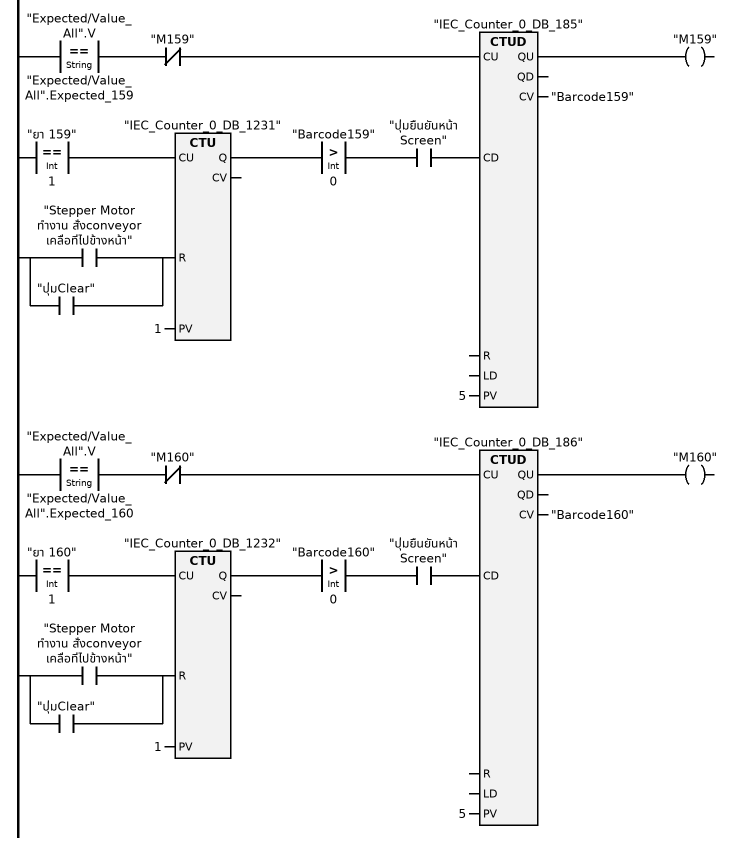
   "IEC_Counter_0_DB_1213".CTU(CU := "ยา 141" = 1,
                           R := "Stepper Motor ทำงาน สั่งconveyor เคลื่อที่ไปข้างหน้า" OR "ปุ่มClear",
                           PV := 1);
   "IEC_Counter_0_DB_167".CTUD(CU := ("Expected/Value_All".V = "Expected/Value_All".Expected_141) AND NOT "M141",
                           CD := "IEC_Counter_0_DB_1213".Q AND ("Barcode141" > 0) AND "ปุ่มยืนยันหน้า Screen",
                           PV := 5,
                           CV => "Barcode141");
   "M141" := "IEC_Counter_0_DB_167".QU;
   "IEC_Counter_0_DB_1214".CTU(CU := "ยา 142" = 1,
                           R := "Stepper Motor ทำงาน สั่งconveyor เคลื่อที่ไปข้างหน้า" OR "ปุ่มClear",
                           PV := 1);
   "IEC_Counter_0_DB_168".CTUD(CU := ("Expected/Value_All".V = "Expected/Value_All".Expected_142) AND NOT "M142",
                           CD := "IEC_Counter_0_DB_1214".Q AND ("Barcode142" > 0) AND "ปุ่มยืนยันหน้า Screen",
                           PV := 5,
                           CV => "Barcode142");
   "M142" := "IEC_Counter_0_DB_168".QU;
   "IEC_Counter_0_DB_1215".CTU(CU := "ยา 143" = 1,
                           R := "Stepper Motor ทำงาน สั่งconveyor เคลื่อที่ไปข้างหน้า" OR "ปุ่มClear",
                           PV := 1);
   "IEC_Counter_0_DB_169".CTUD(CU := ("Expected/Value_All".V = "Expected/Value_All".Expected_143) AND NOT "M143",
                           CD := "IEC_Counter_0_DB_1215".Q AND ("Barcode143" > 0) AND "ปุ่มยืนยันหน้า Screen",
                           PV := 5,
                           CV => "Barcode143");
   "M143" := "IEC_Counter_0_DB_169".QU;
   "IEC_Counter_0_DB_1216".CTU(CU := "ยา 144" = 1,
                           R := "Stepper Motor ทำงาน สั่งconveyor เคลื่อที่ไปข้างหน้า" OR "ปุ่มClear",
                           PV := 1);
   "IEC_Counter_0_DB_170".CTUD(CU := ("Expected/Value_All".V = "Expected/Value_All".Expected_144) AND NOT "M144",
                           CD := "IEC_Counter_0_DB_1216".Q AND ("Barcode144" > 0) AND "ปุ่มยืนยันหน้า Screen",
                           PV := 5,
                           CV => "Barcode144");
   "M144" := "IEC_Counter_0_DB_170".QU;
   "IEC_Counter_0_DB_1217".CTU(CU := "ยา 145" = 1,
                           R := "Stepper Motor ทำงาน สั่งconveyor เคลื่อที่ไปข้างหน้า" OR "ปุ่มClear",
                           PV := 1);
   "IEC_Counter_0_DB_171".CTUD(CU := ("Expected/Value_All".V = "Expected/Value_All".Expected_145) AND NOT "M145",
                           CD := "IEC_Counter_0_DB_1217".Q AND ("Barcode145" > 0) AND "ปุ่มยืนยันหน้า Screen",
                           PV := 5,
                           CV => "Barcode145");
   "M145" := "IEC_Counter_0_DB_171".QU;
   "IEC_Counter_0_DB_1218".CTU(CU := "ยา 146" = 1,
                           R := "Stepper Motor ทำงาน สั่งconveyor เคลื่อที่ไปข้างหน้า" OR "ปุ่มClear",
                           PV := 1);
   "IEC_Counter_0_DB_172".CTUD(CU := ("Expected/Value_All".V = "Expected/Value_All".Expected_146) AND NOT "M146",
                           CD := "IEC_Counter_0_DB_1218".Q AND ("Barcode146" > 0) AND "ปุ่มยืนยันหน้า Screen",
                           PV := 5,
                           CV => "Barcode146");
   "M146" := "IEC_Counter_0_DB_172".QU;
   "IEC_Counter_0_DB_1219".CTU(CU := "ยา 147" = 1,
                           R := "Stepper Motor ทำงาน สั่งconveyor เคลื่อที่ไปข้างหน้า" OR "ปุ่มClear",
                           PV := 1);
   "IEC_Counter_0_DB_173".CTUD(CU := ("Expected/Value_All".V = "Expected/Value_All".Expected_147) AND NOT "M147",
                           CD := "IEC_Counter_0_DB_1219".Q AND ("Barcode147" > 0) AND "ปุ่มยืนยันหน้า Screen",
                           PV := 5,
                           CV => "Barcode147");
   "M147" := "IEC_Counter_0_DB_173".QU;
   "IEC_Counter_0_DB_1220".CTU(CU := "ยา 148" = 1,
                           R := "Stepper Motor ทำงาน สั่งconveyor เคลื่อที่ไปข้างหน้า" OR "ปุ่มClear",
                           PV := 1);
   "IEC_Counter_0_DB_174".CTUD(CU := ("Expected/Value_All".V = "Expected/Value_All".Expected_148) AND NOT "M148",
                           CD := "IEC_Counter_0_DB_1220".Q AND ("Barcode148" > 0) AND "ปุ่มยืนยันหน้า Screen",
                           PV := 5,
                           CV => "Barcode148");
   "M148" := "IEC_Counter_0_DB_174".QU;
   "IEC_Counter_0_DB_1221".CTU(CU := "ยา 149" = 1,
                           R := "Stepper Motor ทำงาน สั่งconveyor เคลื่อที่ไปข้างหน้า" OR "ปุ่มClear",
                           PV := 1);
   "IEC_Counter_0_DB_175".CTUD(CU := ("Expected/Value_All".V = "Expected/Value_All".Expected_149) AND NOT "M149",
                           CD := "IEC_Counter_0_DB_1221".Q AND ("Barcode149" > 0) AND "ปุ่มยืนยันหน้า Screen",
                           PV := 5,
                           CV => "Barcode149");
   "M149" := "IEC_Counter_0_DB_175".QU;
   "IEC_Counter_0_DB_1222".CTU(CU := "ยา 150" = 1,
                           R := "Stepper Motor ทำงาน สั่งconveyor เคลื่อที่ไปข้างหน้า" OR "ปุ่มClear",
                           PV := 1);
   "IEC_Counter_0_DB_176".CTUD(CU := ("Expected/Value_All".V = "Expected/Value_All".Expected_150) AND NOT "M150",
                           CD := "IEC_Counter_0_DB_1222".Q AND ("Barcode150" > 0) AND "ปุ่มยืนยันหน้า Screen",
                           PV := 5,
                           CV => "Barcode150");
   "M150" := "IEC_Counter_0_DB_176".QU;
   "IEC_Counter_0_DB_1223".CTU(CU := "ยา 151" = 1,
                           R := "Stepper Motor ทำงาน สั่งconveyor เคลื่อที่ไปข้างหน้า" OR "ปุ่มClear",
                           PV := 1);
   "IEC_Counter_0_DB_177".CTUD(CU := ("Expected/Value_All".V = "Expected/Value_All".Expected_151) AND NOT "M151",
                           CD := "IEC_Counter_0_DB_1223".Q AND ("Barcode151" > 0) AND "ปุ่มยืนยันหน้า Screen",
                           PV := 5,
                           CV => "Barcode151");
   "M151" := "IEC_Counter_0_DB_177".QU;
   "IEC_Counter_0_DB_1224".CTU(CU := "ยา 152" = 1,
                           R := "Stepper Motor ทำงาน สั่งconveyor เคลื่อที่ไปข้างหน้า" OR "ปุ่มClear",
                           PV := 1);
   "IEC_Counter_0_DB_178".CTUD(CU := ("Expected/Value_All".V = "Expected/Value_All".Expected_152) AND NOT "M152",
                           CD := "IEC_Counter_0_DB_1224".Q AND ("Barcode152" > 0) AND "ปุ่มยืนยันหน้า Screen",
                           PV := 5,
                           CV => "Barcode152");
   "M152" := "IEC_Counter_0_DB_178".QU;
   "IEC_Counter_0_DB_1225".CTU(CU := "ยา 153" = 1,
                           R := "Stepper Motor ทำงาน สั่งconveyor เคลื่อที่ไปข้างหน้า" OR "ปุ่มClear",
                           PV := 1);
   "IEC_Counter_0_DB_179".CTUD(CU := ("Expected/Value_All".V = "Expected/Value_All".Expected_153) AND NOT "M153",
                           CD := "IEC_Counter_0_DB_1225".Q AND ("Barcode153" > 0) AND "ปุ่มยืนยันหน้า Screen",
                           PV := 5,
                           CV => "Barcode153");
   "M153" := "IEC_Counter_0_DB_179".QU;
   "IEC_Counter_0_DB_1226".CTU(CU := "ยา 154" = 1,
                           R := "Stepper Motor ทำงาน สั่งconveyor เคลื่อที่ไปข้างหน้า" OR "ปุ่มClear",
                           PV := 1);
   "IEC_Counter_0_DB_180".CTUD(CU := ("Expected/Value_All".V = "Expected/Value_All".Expected_154) AND NOT "M154",
                           CD := "IEC_Counter_0_DB_1226".Q AND ("Barcode154" > 0) AND "ปุ่มยืนยันหน้า Screen",
                           PV := 5,
                           CV => "Barcode154");
   "M154" := "IEC_Counter_0_DB_180".QU;
   "IEC_Counter_0_DB_1227".CTU(CU := "ยา 155" = 1,
                           R := "Stepper Motor ทำงาน สั่งconveyor เคลื่อที่ไปข้างหน้า" OR "ปุ่มClear",
                           PV := 1);
   "IEC_Counter_0_DB_181".CTUD(CU := ("Expected/Value_All".V = "Expected/Value_All".Expected_155) AND NOT "M155",
                           CD := "IEC_Counter_0_DB_1227".Q AND ("Barcode155" > 0) AND "ปุ่มยืนยันหน้า Screen",
                           PV := 5,
                           CV => "Barcode155");
   "M155" := "IEC_Counter_0_DB_181".QU;
   "IEC_Counter_0_DB_1228".CTU(CU := "ยา 156" = 1,
                           R := "Stepper Motor ทำงาน สั่งconveyor เคลื่อที่ไปข้างหน้า" OR "ปุ่มClear",
                           PV := 1);
   "IEC_Counter_0_DB_182".CTUD(CU := ("Expected/Value_All".V = "Expected/Value_All".Expected_156) AND NOT "M156",
                           CD := "IEC_Counter_0_DB_1228".Q AND ("Barcode156" > 0) AND "ปุ่มยืนยันหน้า Screen",
                           PV := 5,
                           CV => "Barcode156");
   "M156" := "IEC_Counter_0_DB_182".QU;
   "IEC_Counter_0_DB_1229".CTU(CU := "ยา 157" = 1,
                           R := "Stepper Motor ทำงาน สั่งconveyor เคลื่อที่ไปข้างหน้า" OR "ปุ่มClear",
                           PV := 1);
   "IEC_Counter_0_DB_183".CTUD(CU := ("Expected/Value_All".V = "Expected/Value_All".Expected_157) AND NOT "M157",
                           CD := "IEC_Counter_0_DB_1229".Q AND ("Barcode157" > 0) AND "ปุ่มยืนยันหน้า Screen",
                           PV := 5,
                           CV => "Barcode157");
   "M157" := "IEC_Counter_0_DB_183".QU;
   "IEC_Counter_0_DB_1230".CTU(CU := "ยา 158" = 1,
                           R := "Stepper Motor ทำงาน สั่งconveyor เคลื่อที่ไปข้างหน้า" OR "ปุ่มClear",
                           PV := 1);
   "IEC_Counter_0_DB_184".CTUD(CU := ("Expected/Value_All".V = "Expected/Value_All".Expected_158) AND NOT "M158",
                           CD := "IEC_Counter_0_DB_1230".Q AND ("Barcode158" > 0) AND "ปุ่มยืนยันหน้า Screen",
                           PV := 5,
                           CV => "Barcode158");
   "M158" := "IEC_Counter_0_DB_184".QU;
   "IEC_Counter_0_DB_1231".CTU(CU := "ยา 159" = 1,
                           R := "Stepper Motor ทำงาน สั่งconveyor เคลื่อที่ไปข้างหน้า" OR "ปุ่มClear",
                           PV := 1);
   "IEC_Counter_0_DB_185".CTUD(CU := ("Expected/Value_All".V = "Expected/Value_All".Expected_159) AND NOT "M159",
                           CD := "IEC_Counter_0_DB_1231".Q AND ("Barcode159" > 0) AND "ปุ่มยืนยันหน้า Screen",
                           PV := 5,
                           CV => "Barcode159");
   "M159" := "IEC_Counter_0_DB_185".QU;
   "IEC_Counter_0_DB_1232".CTU(CU := "ยา 160" = 1,
                           R := "Stepper Motor ทำงาน สั่งconveyor เคลื่อที่ไปข้างหน้า" OR "ปุ่มClear",
                           PV := 1);
   "IEC_Counter_0_DB_186".CTUD(CU := ("Expected/Value_All".V = "Expected/Value_All".Expected_160) AND NOT "M160",
                           CD := "IEC_Counter_0_DB_1232".Q AND ("Barcode160" > 0) AND "ปุ่มยืนยันหน้า Screen",
                           PV := 5,
                           CV => "Barcode160");
   "M160" := "IEC_Counter_0_DB_186".QU;
END_REGION

REGION Network 9
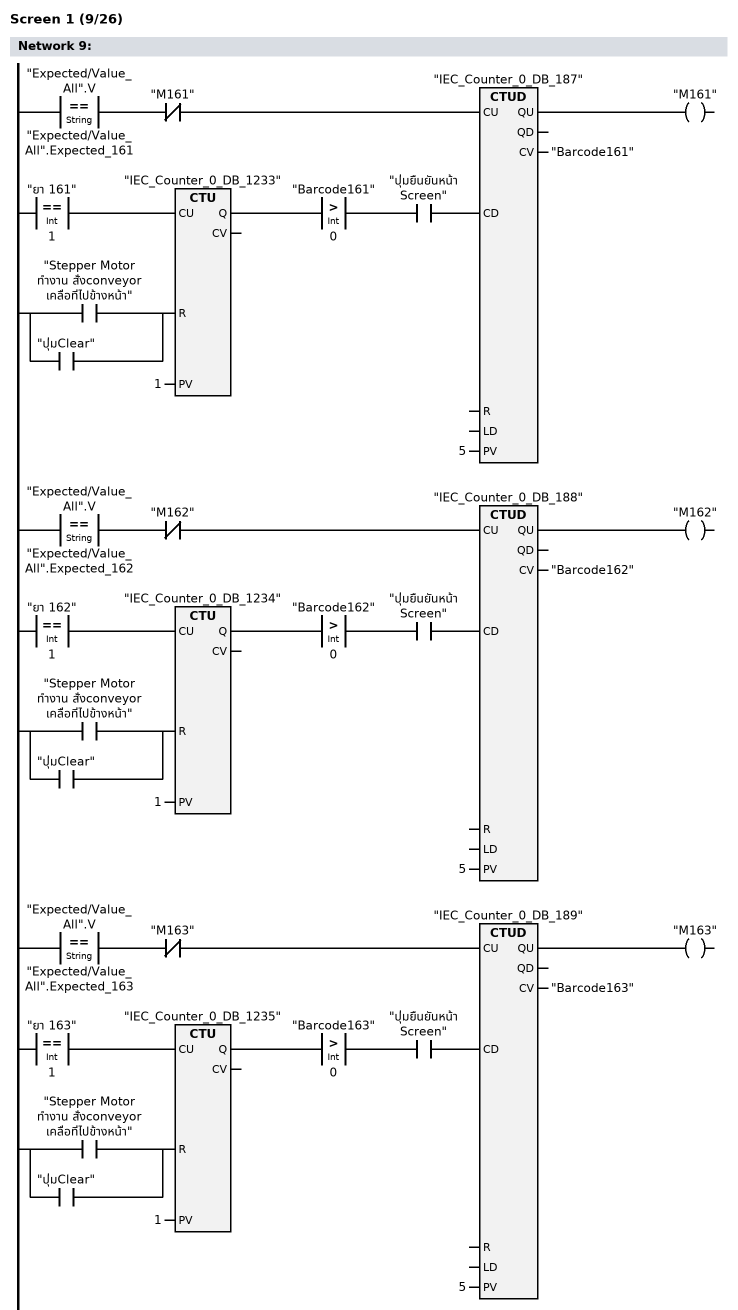
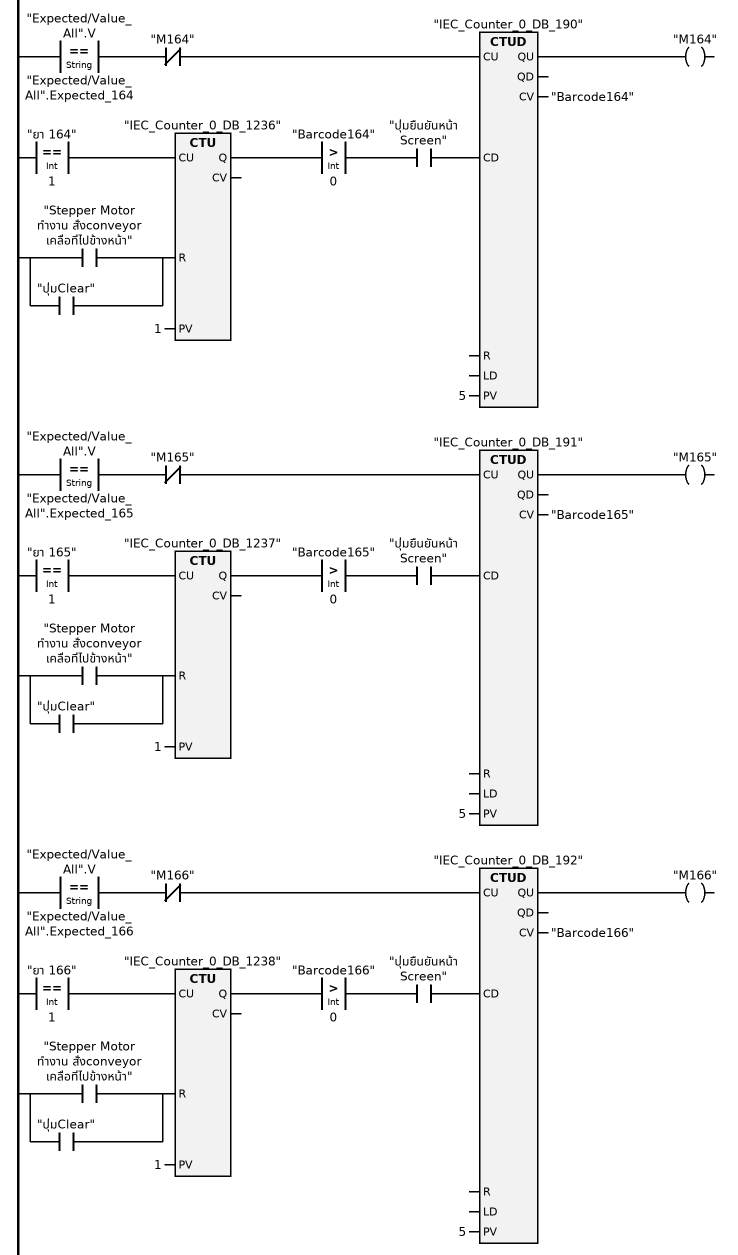
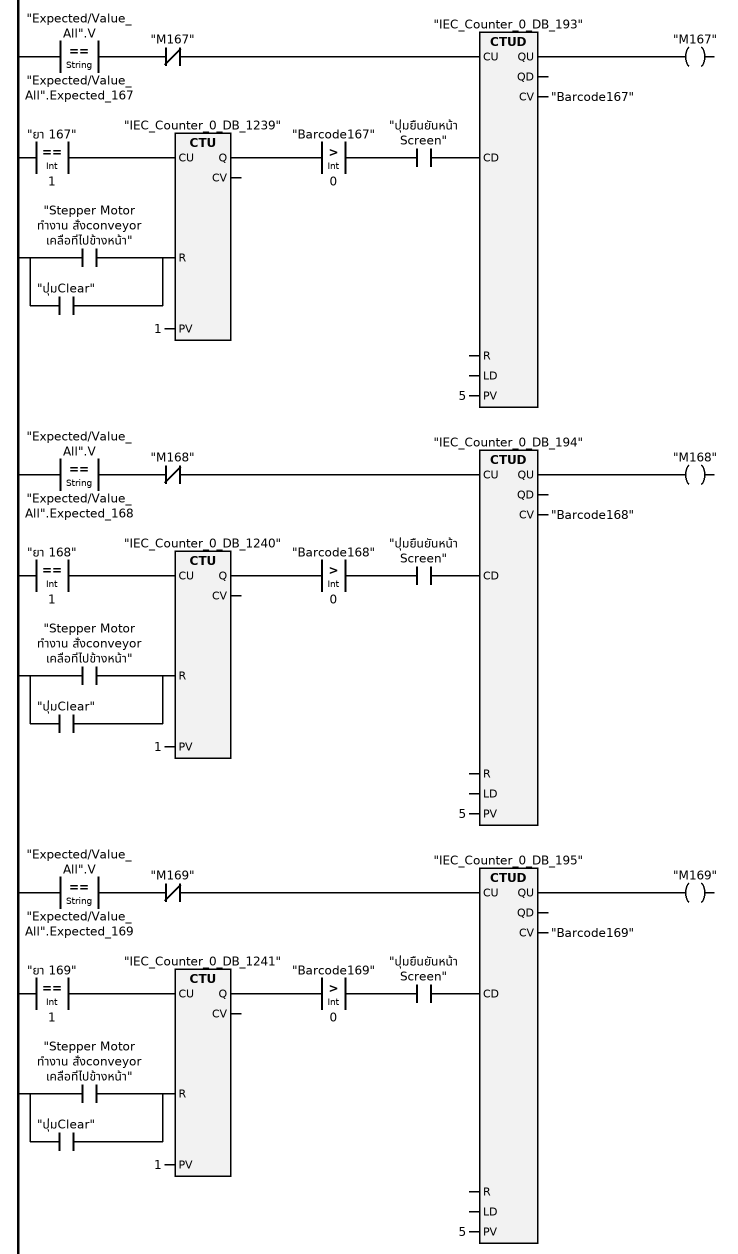
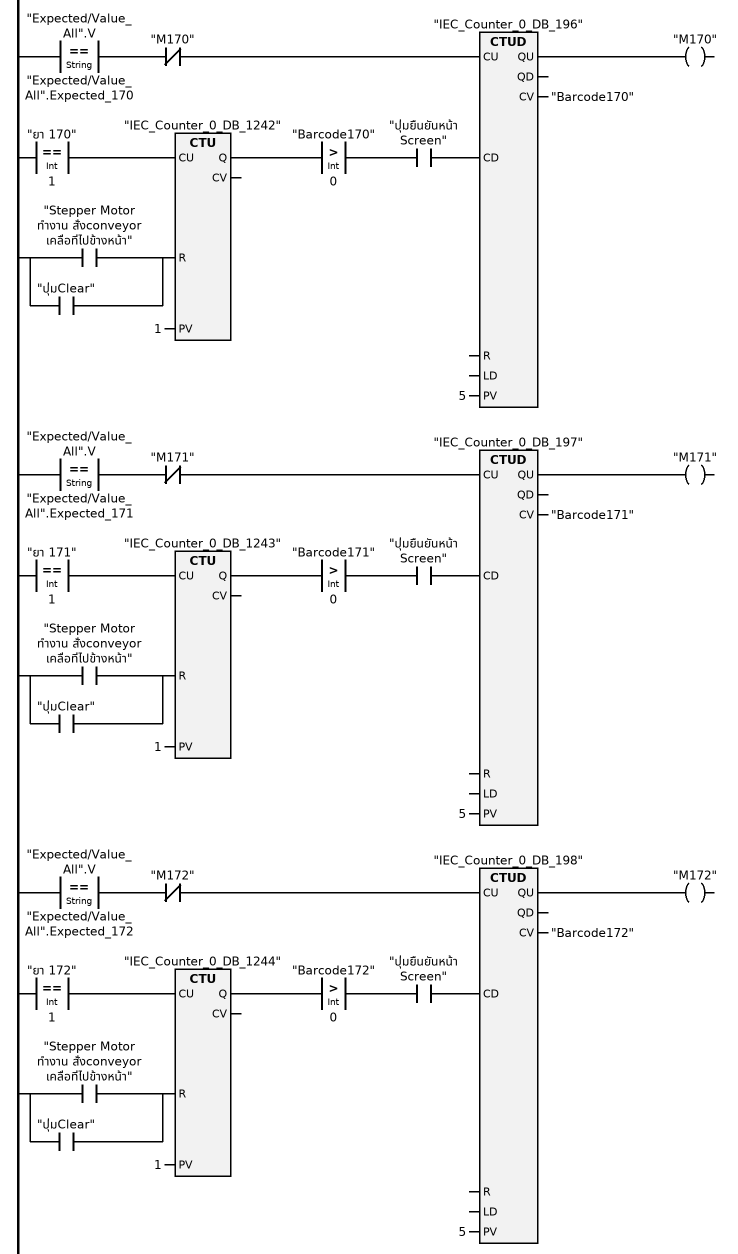
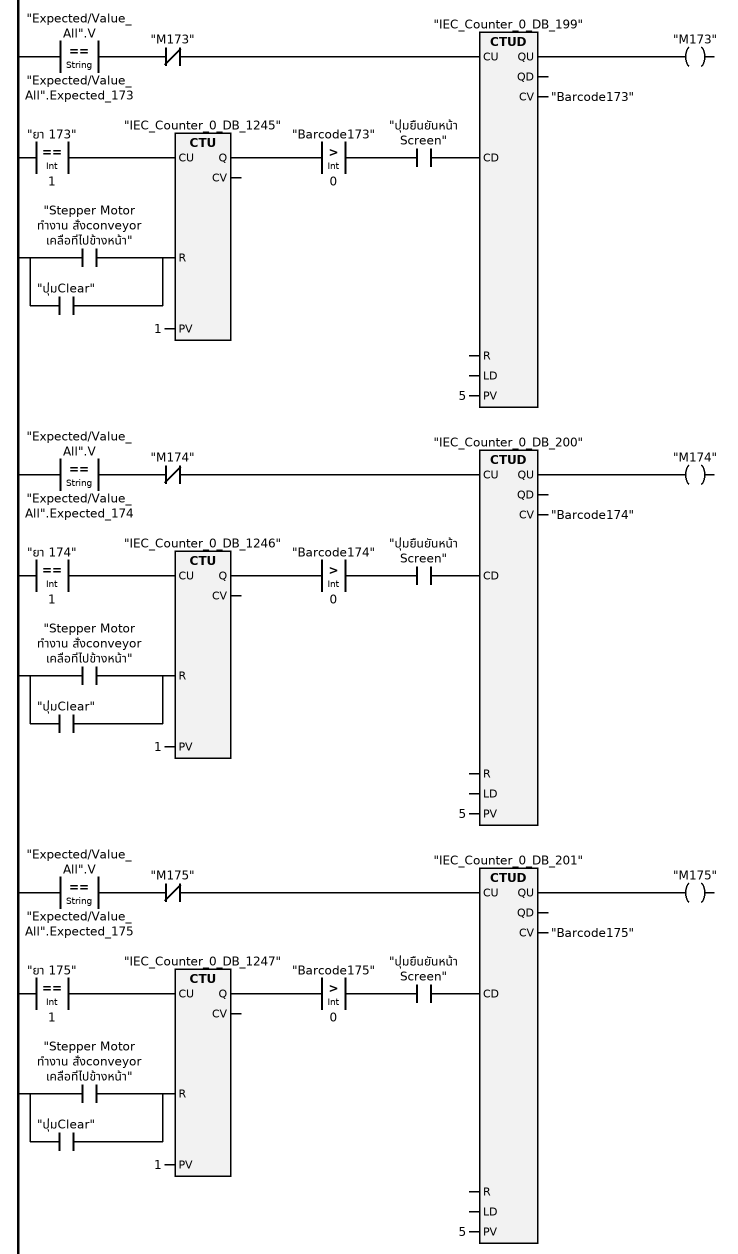
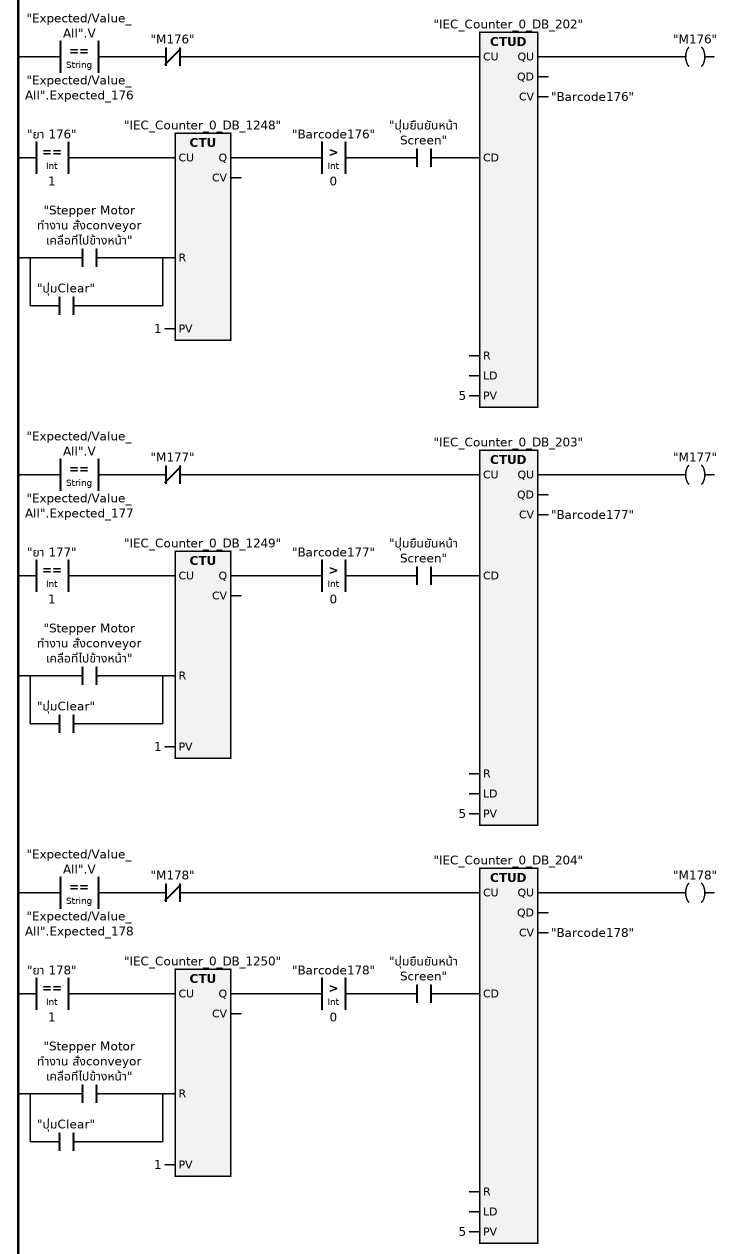
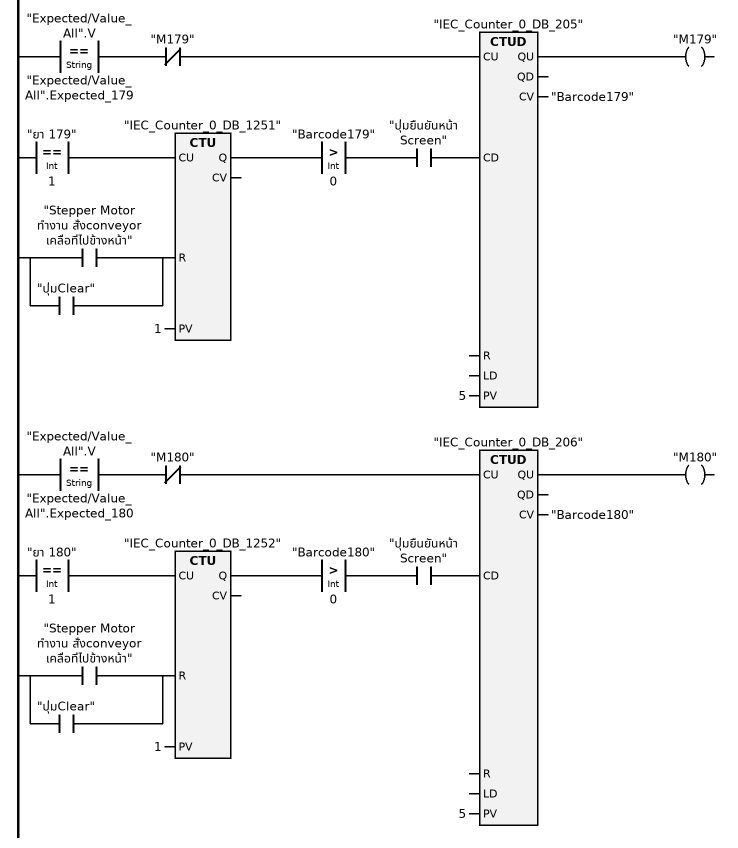
   "IEC_Counter_0_DB_1233".CTU(CU := "ยา 161" = 1,
                           R := "Stepper Motor ทำงาน สั่งconveyor เคลื่อที่ไปข้างหน้า" OR "ปุ่มClear",
                           PV := 1);
   "IEC_Counter_0_DB_187".CTUD(CU := ("Expected/Value_All".V = "Expected/Value_All".Expected_161) AND NOT "M161",
                           CD := "IEC_Counter_0_DB_1233".Q AND ("Barcode161" > 0) AND "ปุ่มยืนยันหน้า Screen",
                           PV := 5,
                           CV => "Barcode161");
   "M161" := "IEC_Counter_0_DB_187".QU;
   "IEC_Counter_0_DB_1234".CTU(CU := "ยา 162" = 1,
                           R := "Stepper Motor ทำงาน สั่งconveyor เคลื่อที่ไปข้างหน้า" OR "ปุ่มClear",
                           PV := 1);
   "IEC_Counter_0_DB_188".CTUD(CU := ("Expected/Value_All".V = "Expected/Value_All".Expected_162) AND NOT "M162",
                           CD := "IEC_Counter_0_DB_1234".Q AND ("Barcode162" > 0) AND "ปุ่มยืนยันหน้า Screen",
                           PV := 5,
                           CV => "Barcode162");
   "M162" := "IEC_Counter_0_DB_188".QU;
   "IEC_Counter_0_DB_1235".CTU(CU := "ยา 163" = 1,
                           R := "Stepper Motor ทำงาน สั่งconveyor เคลื่อที่ไปข้างหน้า" OR "ปุ่มClear",
                           PV := 1);
   "IEC_Counter_0_DB_189".CTUD(CU := ("Expected/Value_All".V = "Expected/Value_All".Expected_163) AND NOT "M163",
                           CD := "IEC_Counter_0_DB_1235".Q AND ("Barcode163" > 0) AND "ปุ่มยืนยันหน้า Screen",
                           PV := 5,
                           CV => "Barcode163");
   "M163" := "IEC_Counter_0_DB_189".QU;
   "IEC_Counter_0_DB_1236".CTU(CU := "ยา 164" = 1,
                           R := "Stepper Motor ทำงาน สั่งconveyor เคลื่อที่ไปข้างหน้า" OR "ปุ่มClear",
                           PV := 1);
   "IEC_Counter_0_DB_190".CTUD(CU := ("Expected/Value_All".V = "Expected/Value_All".Expected_164) AND NOT "M164",
                           CD := "IEC_Counter_0_DB_1236".Q AND ("Barcode164" > 0) AND "ปุ่มยืนยันหน้า Screen",
                           PV := 5,
                           CV => "Barcode164");
   "M164" := "IEC_Counter_0_DB_190".QU;
   "IEC_Counter_0_DB_1237".CTU(CU := "ยา 165" = 1,
                           R := "Stepper Motor ทำงาน สั่งconveyor เคลื่อที่ไปข้างหน้า" OR "ปุ่มClear",
                           PV := 1);
   "IEC_Counter_0_DB_191".CTUD(CU := ("Expected/Value_All".V = "Expected/Value_All".Expected_165) AND NOT "M165",
                           CD := "IEC_Counter_0_DB_1237".Q AND ("Barcode165" > 0) AND "ปุ่มยืนยันหน้า Screen",
                           PV := 5,
                           CV => "Barcode165");
   "M165" := "IEC_Counter_0_DB_191".QU;
   "IEC_Counter_0_DB_1238".CTU(CU := "ยา 166" = 1,
                           R := "Stepper Motor ทำงาน สั่งconveyor เคลื่อที่ไปข้างหน้า" OR "ปุ่มClear",
                           PV := 1);
   "IEC_Counter_0_DB_192".CTUD(CU := ("Expected/Value_All".V = "Expected/Value_All".Expected_166) AND NOT "M166",
                           CD := "IEC_Counter_0_DB_1238".Q AND ("Barcode166" > 0) AND "ปุ่มยืนยันหน้า Screen",
                           PV := 5,
                           CV => "Barcode166");
   "M166" := "IEC_Counter_0_DB_192".QU;
   "IEC_Counter_0_DB_1239".CTU(CU := "ยา 167" = 1,
                           R := "Stepper Motor ทำงาน สั่งconveyor เคลื่อที่ไปข้างหน้า" OR "ปุ่มClear",
                           PV := 1);
   "IEC_Counter_0_DB_193".CTUD(CU := ("Expected/Value_All".V = "Expected/Value_All".Expected_167) AND NOT "M167",
                           CD := "IEC_Counter_0_DB_1239".Q AND ("Barcode167" > 0) AND "ปุ่มยืนยันหน้า Screen",
                           PV := 5,
                           CV => "Barcode167");
   "M167" := "IEC_Counter_0_DB_193".QU;
   "IEC_Counter_0_DB_1240".CTU(CU := "ยา 168" = 1,
                           R := "Stepper Motor ทำงาน สั่งconveyor เคลื่อที่ไปข้างหน้า" OR "ปุ่มClear",
                           PV := 1);
   "IEC_Counter_0_DB_194".CTUD(CU := ("Expected/Value_All".V = "Expected/Value_All".Expected_168) AND NOT "M168",
                           CD := "IEC_Counter_0_DB_1240".Q AND ("Barcode168" > 0) AND "ปุ่มยืนยันหน้า Screen",
                           PV := 5,
                           CV => "Barcode168");
   "M168" := "IEC_Counter_0_DB_194".QU;
   "IEC_Counter_0_DB_1241".CTU(CU := "ยา 169" = 1,
                           R := "Stepper Motor ทำงาน สั่งconveyor เคลื่อที่ไปข้างหน้า" OR "ปุ่มClear",
                           PV := 1);
   "IEC_Counter_0_DB_195".CTUD(CU := ("Expected/Value_All".V = "Expected/Value_All".Expected_169) AND NOT "M169",
                           CD := "IEC_Counter_0_DB_1241".Q AND ("Barcode169" > 0) AND "ปุ่มยืนยันหน้า Screen",
                           PV := 5,
                           CV => "Barcode169");
   "M169" := "IEC_Counter_0_DB_195".QU;
   "IEC_Counter_0_DB_1242".CTU(CU := "ยา 170" = 1,
                           R := "Stepper Motor ทำงาน สั่งconveyor เคลื่อที่ไปข้างหน้า" OR "ปุ่มClear",
                           PV := 1);
   "IEC_Counter_0_DB_196".CTUD(CU := ("Expected/Value_All".V = "Expected/Value_All".Expected_170) AND NOT "M170",
                           CD := "IEC_Counter_0_DB_1242".Q AND ("Barcode170" > 0) AND "ปุ่มยืนยันหน้า Screen",
                           PV := 5,
                           CV => "Barcode170");
   "M170" := "IEC_Counter_0_DB_196".QU;
   "IEC_Counter_0_DB_1243".CTU(CU := "ยา 171" = 1,
                           R := "Stepper Motor ทำงาน สั่งconveyor เคลื่อที่ไปข้างหน้า" OR "ปุ่มClear",
                           PV := 1);
   "IEC_Counter_0_DB_197".CTUD(CU := ("Expected/Value_All".V = "Expected/Value_All".Expected_171) AND NOT "M171",
                           CD := "IEC_Counter_0_DB_1243".Q AND ("Barcode171" > 0) AND "ปุ่มยืนยันหน้า Screen",
                           PV := 5,
                           CV => "Barcode171");
   "M171" := "IEC_Counter_0_DB_197".QU;
   "IEC_Counter_0_DB_1244".CTU(CU := "ยา 172" = 1,
                           R := "Stepper Motor ทำงาน สั่งconveyor เคลื่อที่ไปข้างหน้า" OR "ปุ่มClear",
                           PV := 1);
   "IEC_Counter_0_DB_198".CTUD(CU := ("Expected/Value_All".V = "Expected/Value_All".Expected_172) AND NOT "M172",
                           CD := "IEC_Counter_0_DB_1244".Q AND ("Barcode172" > 0) AND "ปุ่มยืนยันหน้า Screen",
                           PV := 5,
                           CV => "Barcode172");
   "M172" := "IEC_Counter_0_DB_198".QU;
   "IEC_Counter_0_DB_1245".CTU(CU := "ยา 173" = 1,
                           R := "Stepper Motor ทำงาน สั่งconveyor เคลื่อที่ไปข้างหน้า" OR "ปุ่มClear",
                           PV := 1);
   "IEC_Counter_0_DB_199".CTUD(CU := ("Expected/Value_All".V = "Expected/Value_All".Expected_173) AND NOT "M173",
                           CD := "IEC_Counter_0_DB_1245".Q AND ("Barcode173" > 0) AND "ปุ่มยืนยันหน้า Screen",
                           PV := 5,
                           CV => "Barcode173");
   "M173" := "IEC_Counter_0_DB_199".QU;
   "IEC_Counter_0_DB_1246".CTU(CU := "ยา 174" = 1,
                           R := "Stepper Motor ทำงาน สั่งconveyor เคลื่อที่ไปข้างหน้า" OR "ปุ่มClear",
                           PV := 1);
   "IEC_Counter_0_DB_200".CTUD(CU := ("Expected/Value_All".V = "Expected/Value_All".Expected_174) AND NOT "M174",
                           CD := "IEC_Counter_0_DB_1246".Q AND ("Barcode174" > 0) AND "ปุ่มยืนยันหน้า Screen",
                           PV := 5,
                           CV => "Barcode174");
   "M174" := "IEC_Counter_0_DB_200".QU;
   "IEC_Counter_0_DB_1247".CTU(CU := "ยา 175" = 1,
                           R := "Stepper Motor ทำงาน สั่งconveyor เคลื่อที่ไปข้างหน้า" OR "ปุ่มClear",
                           PV := 1);
   "IEC_Counter_0_DB_201".CTUD(CU := ("Expected/Value_All".V = "Expected/Value_All".Expected_175) AND NOT "M175",
                           CD := "IEC_Counter_0_DB_1247".Q AND ("Barcode175" > 0) AND "ปุ่มยืนยันหน้า Screen",
                           PV := 5,
                           CV => "Barcode175");
   "M175" := "IEC_Counter_0_DB_201".QU;
   "IEC_Counter_0_DB_1248".CTU(CU := "ยา 176" = 1,
                           R := "Stepper Motor ทำงาน สั่งconveyor เคลื่อที่ไปข้างหน้า" OR "ปุ่มClear",
                           PV := 1);
   "IEC_Counter_0_DB_202".CTUD(CU := ("Expected/Value_All".V = "Expected/Value_All".Expected_176) AND NOT "M176",
                           CD := "IEC_Counter_0_DB_1248".Q AND ("Barcode176" > 0) AND "ปุ่มยืนยันหน้า Screen",
                           PV := 5,
                           CV => "Barcode176");
   "M176" := "IEC_Counter_0_DB_202".QU;
   "IEC_Counter_0_DB_1249".CTU(CU := "ยา 177" = 1,
                           R := "Stepper Motor ทำงาน สั่งconveyor เคลื่อที่ไปข้างหน้า" OR "ปุ่มClear",
                           PV := 1);
   "IEC_Counter_0_DB_203".CTUD(CU := ("Expected/Value_All".V = "Expected/Value_All".Expected_177) AND NOT "M177",
                           CD := "IEC_Counter_0_DB_1249".Q AND ("Barcode177" > 0) AND "ปุ่มยืนยันหน้า Screen",
                           PV := 5,
                           CV => "Barcode177");
   "M177" := "IEC_Counter_0_DB_203".QU;
   "IEC_Counter_0_DB_1250".CTU(CU := "ยา 178" = 1,
                           R := "Stepper Motor ทำงาน สั่งconveyor เคลื่อที่ไปข้างหน้า" OR "ปุ่มClear",
                           PV := 1);
   "IEC_Counter_0_DB_204".CTUD(CU := ("Expected/Value_All".V = "Expected/Value_All".Expected_178) AND NOT "M178",
                           CD := "IEC_Counter_0_DB_1250".Q AND ("Barcode178" > 0) AND "ปุ่มยืนยันหน้า Screen",
                           PV := 5,
                           CV => "Barcode178");
   "M178" := "IEC_Counter_0_DB_204".QU;
   "IEC_Counter_0_DB_1251".CTU(CU := "ยา 179" = 1,
                           R := "Stepper Motor ทำงาน สั่งconveyor เคลื่อที่ไปข้างหน้า" OR "ปุ่มClear",
                           PV := 1);
   "IEC_Counter_0_DB_205".CTUD(CU := ("Expected/Value_All".V = "Expected/Value_All".Expected_179) AND NOT "M179",
                           CD := "IEC_Counter_0_DB_1251".Q AND ("Barcode179" > 0) AND "ปุ่มยืนยันหน้า Screen",
                           PV := 5,
                           CV => "Barcode179");
   "M179" := "IEC_Counter_0_DB_205".QU;
   "IEC_Counter_0_DB_1252".CTU(CU := "ยา 180" = 1,
                           R := "Stepper Motor ทำงาน สั่งconveyor เคลื่อที่ไปข้างหน้า" OR "ปุ่มClear",
                           PV := 1);
   "IEC_Counter_0_DB_206".CTUD(CU := ("Expected/Value_All".V = "Expected/Value_All".Expected_180) AND NOT "M180",
                           CD := "IEC_Counter_0_DB_1252".Q AND ("Barcode180" > 0) AND "ปุ่มยืนยันหน้า Screen",
                           PV := 5,
                           CV => "Barcode180");
   "M180" := "IEC_Counter_0_DB_206".QU;
END_REGION

REGION Network 10
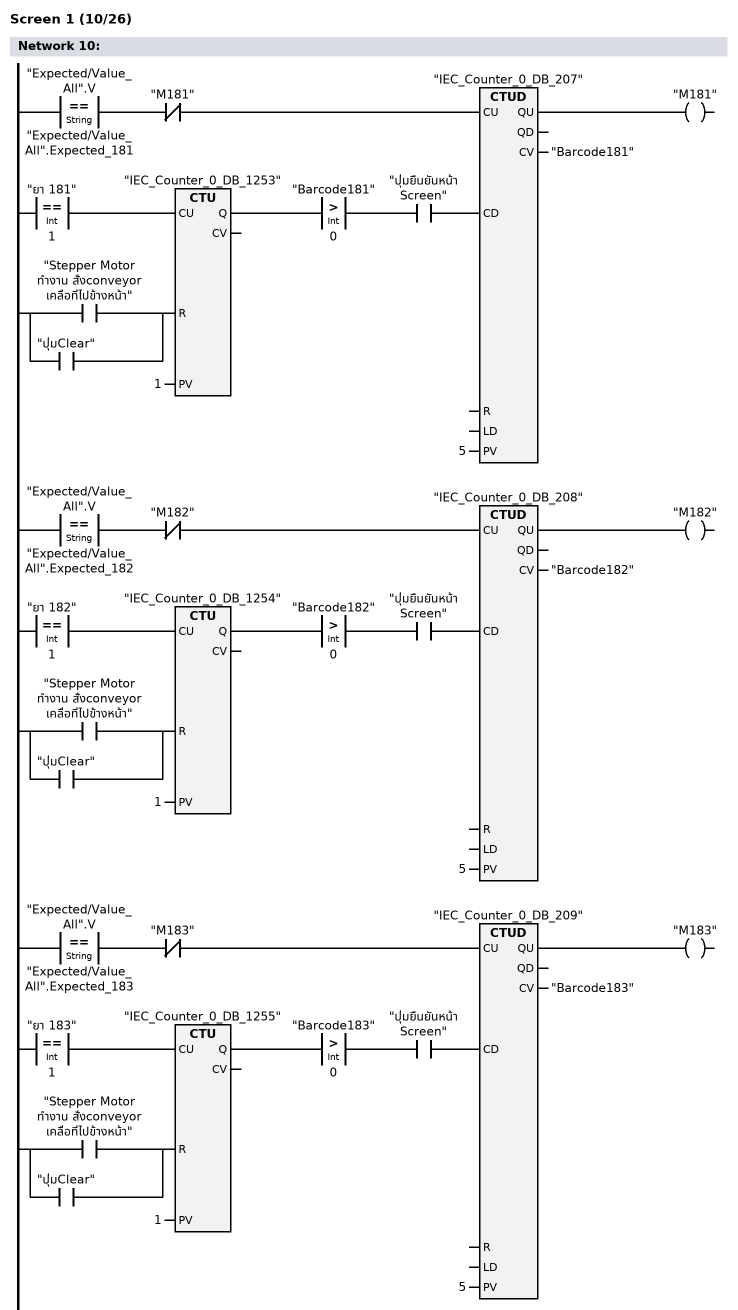
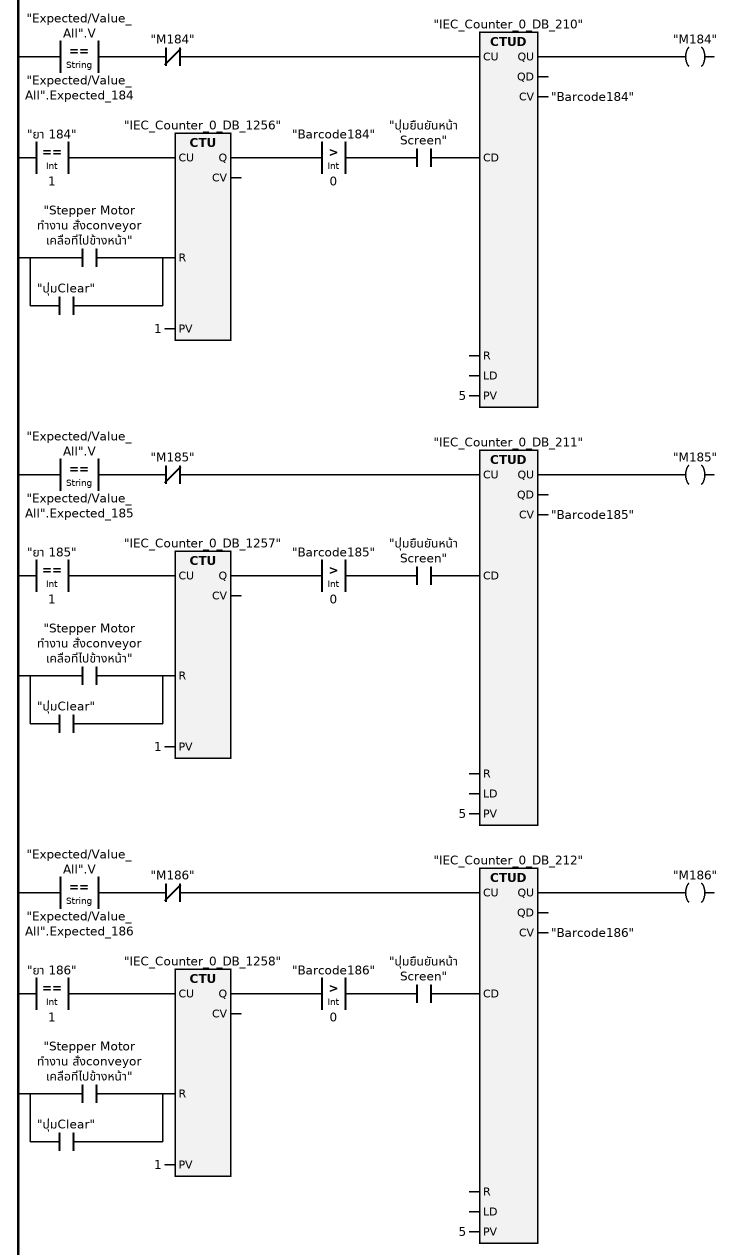
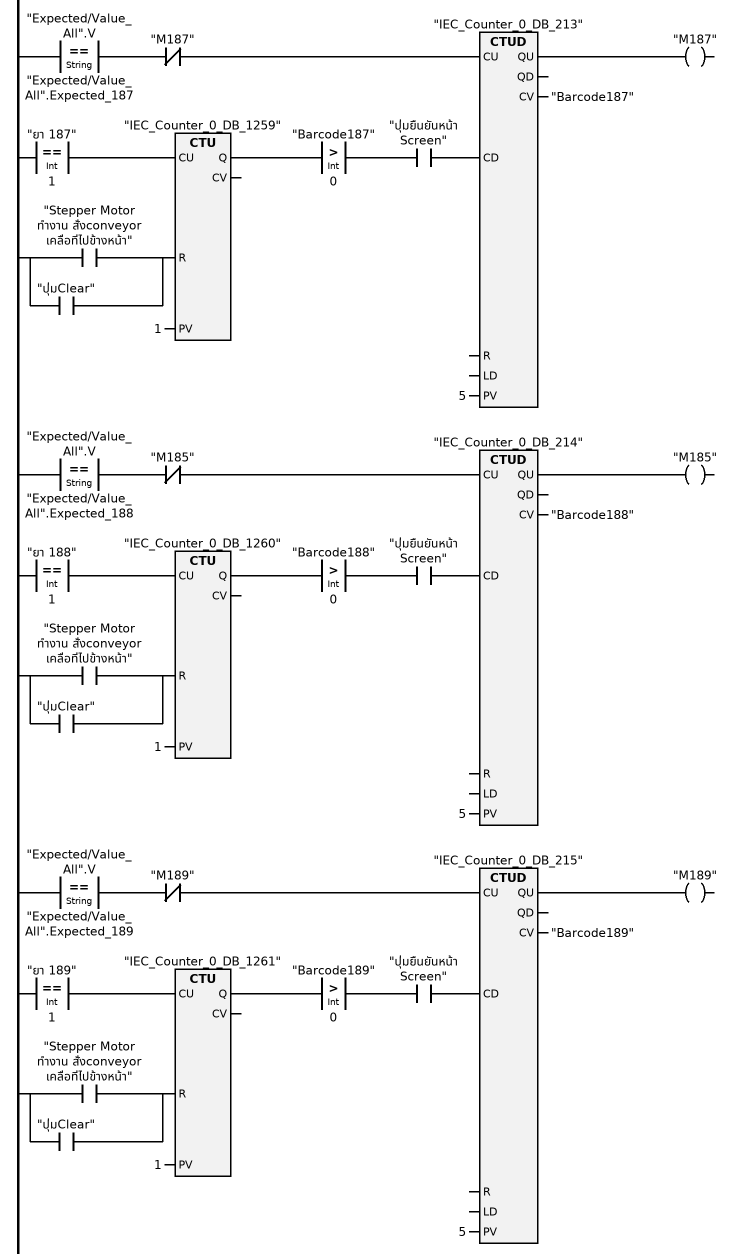
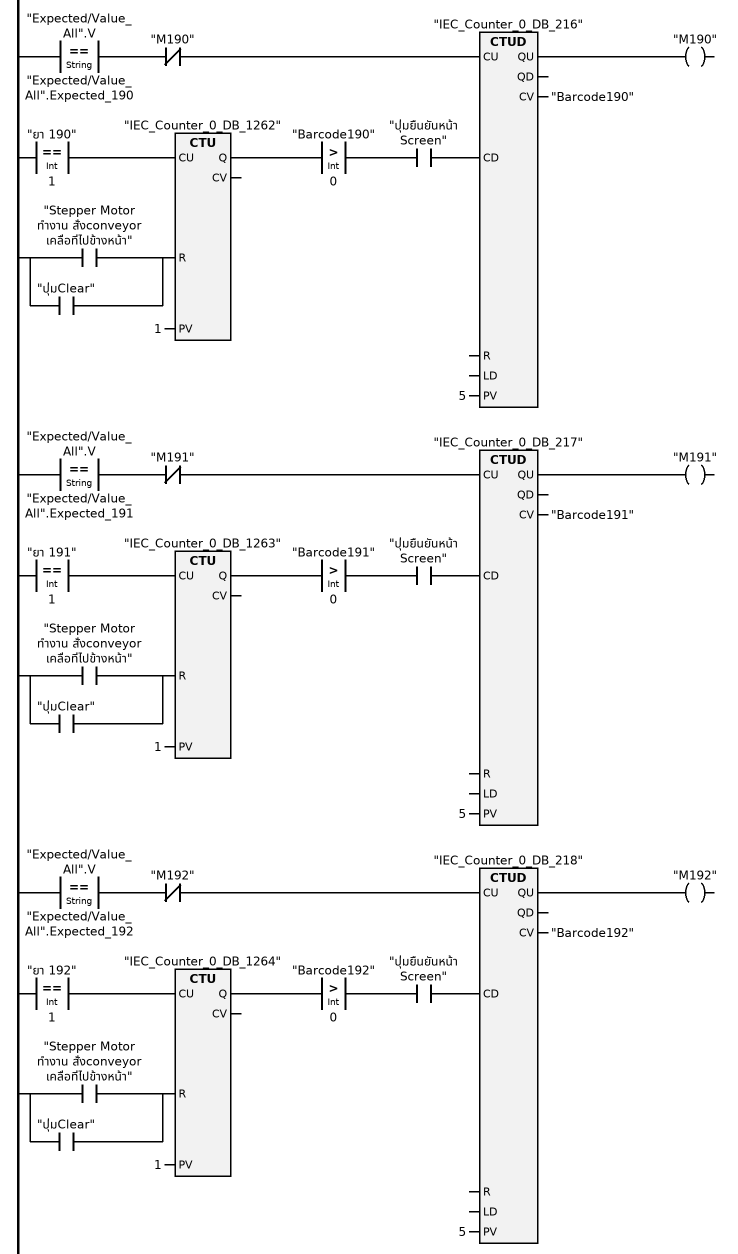
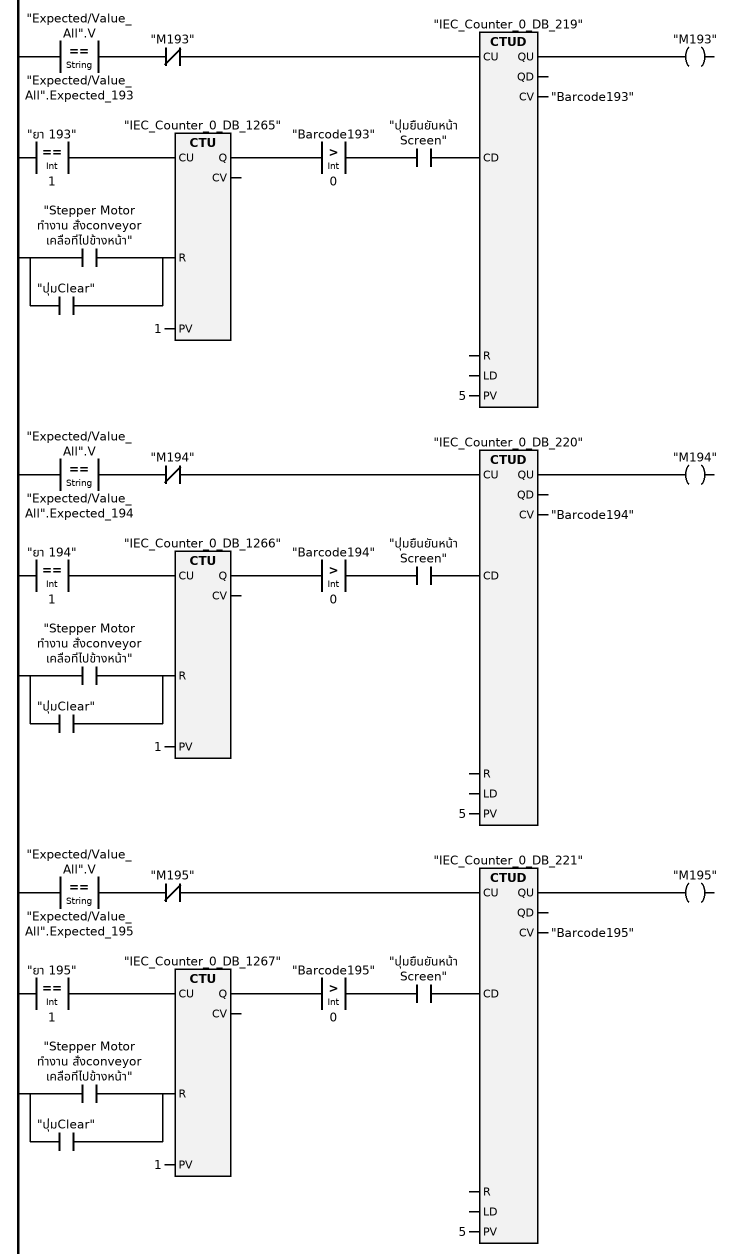
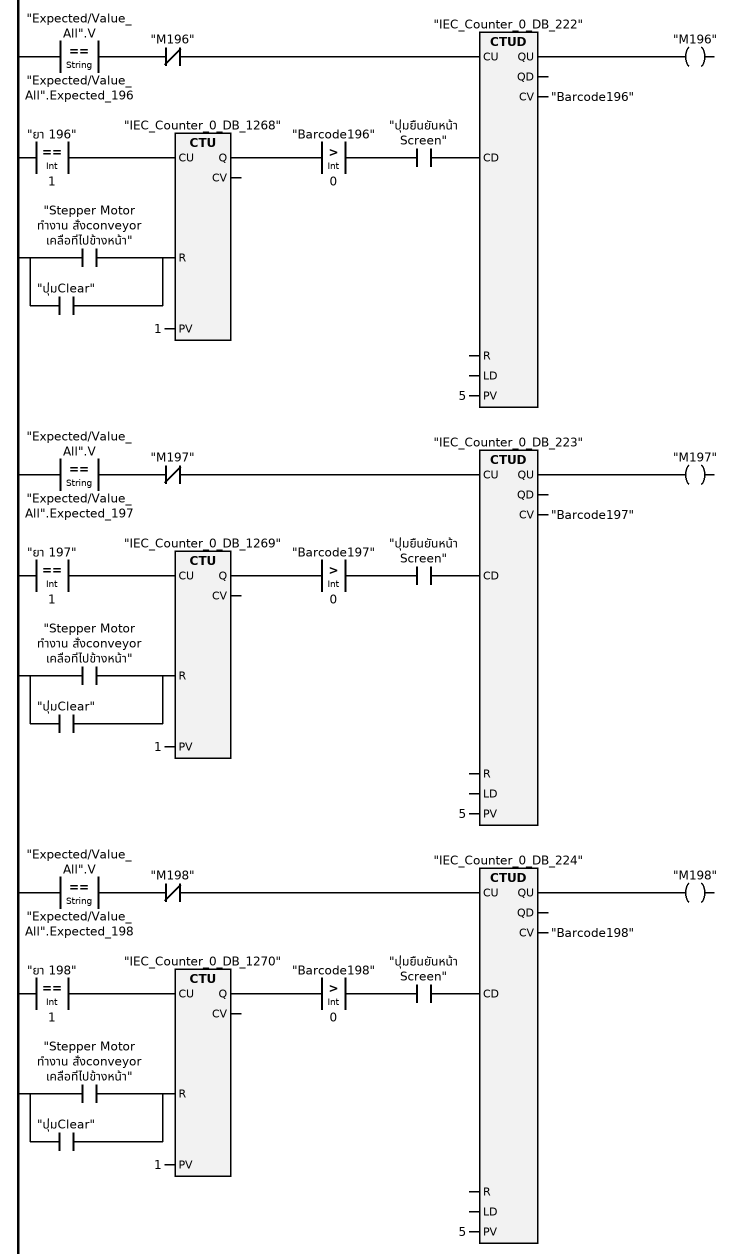
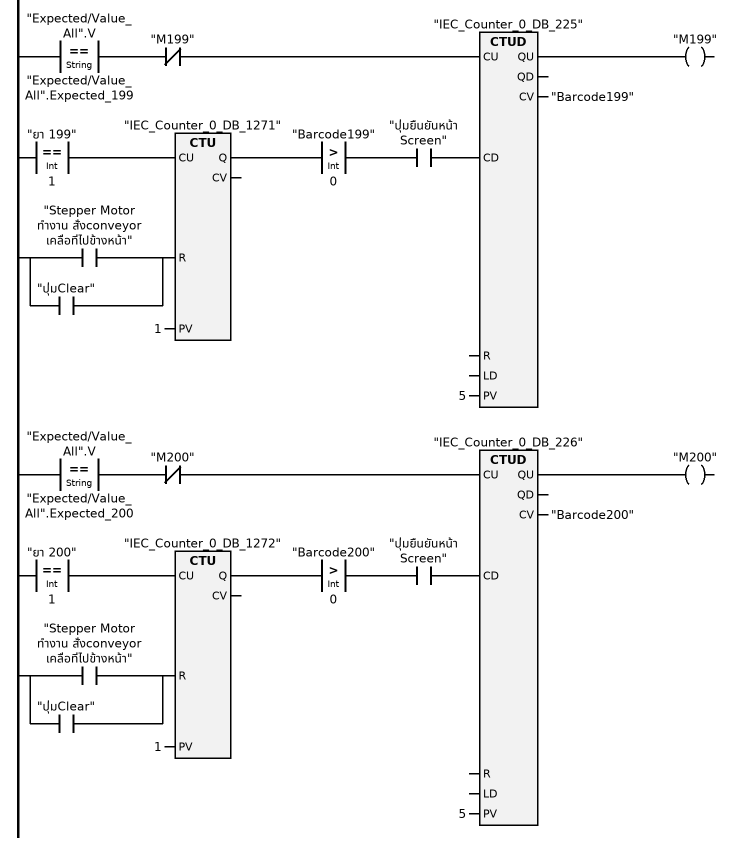
   "IEC_Counter_0_DB_1253".CTU(CU := "ยา 181" = 1,
                           R := "Stepper Motor ทำงาน สั่งconveyor เคลื่อที่ไปข้างหน้า" OR "ปุ่มClear",
                           PV := 1);
   "IEC_Counter_0_DB_207".CTUD(CU := ("Expected/Value_All".V = "Expected/Value_All".Expected_181) AND NOT "M181",
                           CD := "IEC_Counter_0_DB_1253".Q AND ("Barcode181" > 0) AND "ปุ่มยืนยันหน้า Screen",
                           PV := 5,
                           CV => "Barcode181");
   "M181" := "IEC_Counter_0_DB_207".QU;
   "IEC_Counter_0_DB_1254".CTU(CU := "ยา 182" = 1,
                           R := "Stepper Motor ทำงาน สั่งconveyor เคลื่อที่ไปข้างหน้า" OR "ปุ่มClear",
                           PV := 1);
   "IEC_Counter_0_DB_208".CTUD(CU := ("Expected/Value_All".V = "Expected/Value_All".Expected_182) AND NOT "M182",
                           CD := "IEC_Counter_0_DB_1254".Q AND ("Barcode182" > 0) AND "ปุ่มยืนยันหน้า Screen",
                           PV := 5,
                           CV => "Barcode182");
   "M182" := "IEC_Counter_0_DB_208".QU;
   "IEC_Counter_0_DB_1255".CTU(CU := "ยา 183" = 1,
                           R := "Stepper Motor ทำงาน สั่งconveyor เคลื่อที่ไปข้างหน้า" OR "ปุ่มClear",
                           PV := 1);
   "IEC_Counter_0_DB_209".CTUD(CU := ("Expected/Value_All".V = "Expected/Value_All".Expected_183) AND NOT "M183",
                           CD := "IEC_Counter_0_DB_1255".Q AND ("Barcode183" > 0) AND "ปุ่มยืนยันหน้า Screen",
                           PV := 5,
                           CV => "Barcode183");
   "M183" := "IEC_Counter_0_DB_209".QU;
   "IEC_Counter_0_DB_1256".CTU(CU := "ยา 184" = 1,
                           R := "Stepper Motor ทำงาน สั่งconveyor เคลื่อที่ไปข้างหน้า" OR "ปุ่มClear",
                           PV := 1);
   "IEC_Counter_0_DB_210".CTUD(CU := ("Expected/Value_All".V = "Expected/Value_All".Expected_184) AND NOT "M184",
                           CD := "IEC_Counter_0_DB_1256".Q AND ("Barcode184" > 0) AND "ปุ่มยืนยันหน้า Screen",
                           PV := 5,
                           CV => "Barcode184");
   "M184" := "IEC_Counter_0_DB_210".QU;
   "IEC_Counter_0_DB_1257".CTU(CU := "ยา 185" = 1,
                           R := "Stepper Motor ทำงาน สั่งconveyor เคลื่อที่ไปข้างหน้า" OR "ปุ่มClear",
                           PV := 1);
   "IEC_Counter_0_DB_211".CTUD(CU := ("Expected/Value_All".V = "Expected/Value_All".Expected_185) AND NOT "M185",
                           CD := "IEC_Counter_0_DB_1257".Q AND ("Barcode185" > 0) AND "ปุ่มยืนยันหน้า Screen",
                           PV := 5,
                           CV => "Barcode185");
   "M185" := "IEC_Counter_0_DB_211".QU;
   "IEC_Counter_0_DB_1258".CTU(CU := "ยา 186" = 1,
                           R := "Stepper Motor ทำงาน สั่งconveyor เคลื่อที่ไปข้างหน้า" OR "ปุ่มClear",
                           PV := 1);
   "IEC_Counter_0_DB_212".CTUD(CU := ("Expected/Value_All".V = "Expected/Value_All".Expected_186) AND NOT "M186",
                           CD := "IEC_Counter_0_DB_1258".Q AND ("Barcode186" > 0) AND "ปุ่มยืนยันหน้า Screen",
                           PV := 5,
                           CV => "Barcode186");
   "M186" := "IEC_Counter_0_DB_212".QU;
   "IEC_Counter_0_DB_1259".CTU(CU := "ยา 187" = 1,
                           R := "Stepper Motor ทำงาน สั่งconveyor เคลื่อที่ไปข้างหน้า" OR "ปุ่มClear",
                           PV := 1);
   "IEC_Counter_0_DB_213".CTUD(CU := ("Expected/Value_All".V = "Expected/Value_All".Expected_187) AND NOT "M187",
                           CD := "IEC_Counter_0_DB_1259".Q AND ("Barcode187" > 0) AND "ปุ่มยืนยันหน้า Screen",
                           PV := 5,
                           CV => "Barcode187");
   "M187" := "IEC_Counter_0_DB_213".QU;
   "IEC_Counter_0_DB_1260".CTU(CU := "ยา 188" = 1,
                           R := "Stepper Motor ทำงาน สั่งconveyor เคลื่อที่ไปข้างหน้า" OR "ปุ่มClear",
                           PV := 1);
   "IEC_Counter_0_DB_214".CTUD(CU := ("Expected/Value_All".V = "Expected/Value_All".Expected_188) AND NOT "M185",
                           CD := "IEC_Counter_0_DB_1260".Q AND ("Barcode188" > 0) AND "ปุ่มยืนยันหน้า Screen",
                           PV := 5,
                           CV => "Barcode188");
   "M185" := "IEC_Counter_0_DB_214".QU;
   "IEC_Counter_0_DB_1261".CTU(CU := "ยา 189" = 1,
                           R := "Stepper Motor ทำงาน สั่งconveyor เคลื่อที่ไปข้างหน้า" OR "ปุ่มClear",
                           PV := 1);
   "IEC_Counter_0_DB_215".CTUD(CU := ("Expected/Value_All".V = "Expected/Value_All".Expected_189) AND NOT "M189",
                           CD := "IEC_Counter_0_DB_1261".Q AND ("Barcode189" > 0) AND "ปุ่มยืนยันหน้า Screen",
                           PV := 5,
                           CV => "Barcode189");
   "M189" := "IEC_Counter_0_DB_215".QU;
   "IEC_Counter_0_DB_1262".CTU(CU := "ยา 190" = 1,
                           R := "Stepper Motor ทำงาน สั่งconveyor เคลื่อที่ไปข้างหน้า" OR "ปุ่มClear",
                           PV := 1);
   "IEC_Counter_0_DB_216".CTUD(CU := ("Expected/Value_All".V = "Expected/Value_All".Expected_190) AND NOT "M190",
                           CD := "IEC_Counter_0_DB_1262".Q AND ("Barcode190" > 0) AND "ปุ่มยืนยันหน้า Screen",
                           PV := 5,
                           CV => "Barcode190");
   "M190" := "IEC_Counter_0_DB_216".QU;
   "IEC_Counter_0_DB_1263".CTU(CU := "ยา 191" = 1,
                           R := "Stepper Motor ทำงาน สั่งconveyor เคลื่อที่ไปข้างหน้า" OR "ปุ่มClear",
                           PV := 1);
   "IEC_Counter_0_DB_217".CTUD(CU := ("Expected/Value_All".V = "Expected/Value_All".Expected_191) AND NOT "M191",
                           CD := "IEC_Counter_0_DB_1263".Q AND ("Barcode191" > 0) AND "ปุ่มยืนยันหน้า Screen",
                           PV := 5,
                           CV => "Barcode191");
   "M191" := "IEC_Counter_0_DB_217".QU;
   "IEC_Counter_0_DB_1264".CTU(CU := "ยา 192" = 1,
                           R := "Stepper Motor ทำงาน สั่งconveyor เคลื่อที่ไปข้างหน้า" OR "ปุ่มClear",
                           PV := 1);
   "IEC_Counter_0_DB_218".CTUD(CU := ("Expected/Value_All".V = "Expected/Value_All".Expected_192) AND NOT "M192",
                           CD := "IEC_Counter_0_DB_1264".Q AND ("Barcode192" > 0) AND "ปุ่มยืนยันหน้า Screen",
                           PV := 5,
                           CV => "Barcode192");
   "M192" := "IEC_Counter_0_DB_218".QU;
   "IEC_Counter_0_DB_1265".CTU(CU := "ยา 193" = 1,
                           R := "Stepper Motor ทำงาน สั่งconveyor เคลื่อที่ไปข้างหน้า" OR "ปุ่มClear",
                           PV := 1);
   "IEC_Counter_0_DB_219".CTUD(CU := ("Expected/Value_All".V = "Expected/Value_All".Expected_193) AND NOT "M193",
                           CD := "IEC_Counter_0_DB_1265".Q AND ("Barcode193" > 0) AND "ปุ่มยืนยันหน้า Screen",
                           PV := 5,
                           CV => "Barcode193");
   "M193" := "IEC_Counter_0_DB_219".QU;
   "IEC_Counter_0_DB_1266".CTU(CU := "ยา 194" = 1,
                           R := "Stepper Motor ทำงาน สั่งconveyor เคลื่อที่ไปข้างหน้า" OR "ปุ่มClear",
                           PV := 1);
   "IEC_Counter_0_DB_220".CTUD(CU := ("Expected/Value_All".V = "Expected/Value_All".Expected_194) AND NOT "M194",
                           CD := "IEC_Counter_0_DB_1266".Q AND ("Barcode194" > 0) AND "ปุ่มยืนยันหน้า Screen",
                           PV := 5,
                           CV => "Barcode194");
   "M194" := "IEC_Counter_0_DB_220".QU;
   "IEC_Counter_0_DB_1267".CTU(CU := "ยา 195" = 1,
                           R := "Stepper Motor ทำงาน สั่งconveyor เคลื่อที่ไปข้างหน้า" OR "ปุ่มClear",
                           PV := 1);
   "IEC_Counter_0_DB_221".CTUD(CU := ("Expected/Value_All".V = "Expected/Value_All".Expected_195) AND NOT "M195",
                           CD := "IEC_Counter_0_DB_1267".Q AND ("Barcode195" > 0) AND "ปุ่มยืนยันหน้า Screen",
                           PV := 5,
                           CV => "Barcode195");
   "M195" := "IEC_Counter_0_DB_221".QU;
   "IEC_Counter_0_DB_1268".CTU(CU := "ยา 196" = 1,
                           R := "Stepper Motor ทำงาน สั่งconveyor เคลื่อที่ไปข้างหน้า" OR "ปุ่มClear",
                           PV := 1);
   "IEC_Counter_0_DB_222".CTUD(CU := ("Expected/Value_All".V = "Expected/Value_All".Expected_196) AND NOT "M196",
                           CD := "IEC_Counter_0_DB_1268".Q AND ("Barcode196" > 0) AND "ปุ่มยืนยันหน้า Screen",
                           PV := 5,
                           CV => "Barcode196");
   "M196" := "IEC_Counter_0_DB_222".QU;
   "IEC_Counter_0_DB_1269".CTU(CU := "ยา 197" = 1,
                           R := "Stepper Motor ทำงาน สั่งconveyor เคลื่อที่ไปข้างหน้า" OR "ปุ่มClear",
                           PV := 1);
   "IEC_Counter_0_DB_223".CTUD(CU := ("Expected/Value_All".V = "Expected/Value_All".Expected_197) AND NOT "M197",
                           CD := "IEC_Counter_0_DB_1269".Q AND ("Barcode197" > 0) AND "ปุ่มยืนยันหน้า Screen",
                           PV := 5,
                           CV => "Barcode197");
   "M197" := "IEC_Counter_0_DB_223".QU;
   "IEC_Counter_0_DB_1270".CTU(CU := "ยา 198" = 1,
                           R := "Stepper Motor ทำงาน สั่งconveyor เคลื่อที่ไปข้างหน้า" OR "ปุ่มClear",
                           PV := 1);
   "IEC_Counter_0_DB_224".CTUD(CU := ("Expected/Value_All".V = "Expected/Value_All".Expected_198) AND NOT "M198",
                           CD := "IEC_Counter_0_DB_1270".Q AND ("Barcode198" > 0) AND "ปุ่มยืนยันหน้า Screen",
                           PV := 5,
                           CV => "Barcode198");
   "M198" := "IEC_Counter_0_DB_224".QU;
   "IEC_Counter_0_DB_1271".CTU(CU := "ยา 199" = 1,
                           R := "Stepper Motor ทำงาน สั่งconveyor เคลื่อที่ไปข้างหน้า" OR "ปุ่มClear",
                           PV := 1);
   "IEC_Counter_0_DB_225".CTUD(CU := ("Expected/Value_All".V = "Expected/Value_All".Expected_199) AND NOT "M199",
                           CD := "IEC_Counter_0_DB_1271".Q AND ("Barcode199" > 0) AND "ปุ่มยืนยันหน้า Screen",
                           PV := 5,
                           CV => "Barcode199");
   "M199" := "IEC_Counter_0_DB_225".QU;
   "IEC_Counter_0_DB_1272".CTU(CU := "ยา 200" = 1,
                           R := "Stepper Motor ทำงาน สั่งconveyor เคลื่อที่ไปข้างหน้า" OR "ปุ่มClear",
                           PV := 1);
   "IEC_Counter_0_DB_226".CTUD(CU := ("Expected/Value_All".V = "Expected/Value_All".Expected_200) AND NOT "M200",
                           CD := "IEC_Counter_0_DB_1272".Q AND ("Barcode200" > 0) AND "ปุ่มยืนยันหน้า Screen",
                           PV := 5,
                           CV => "Barcode200");
   "M200" := "IEC_Counter_0_DB_226".QU;
END_REGION

REGION Network 11
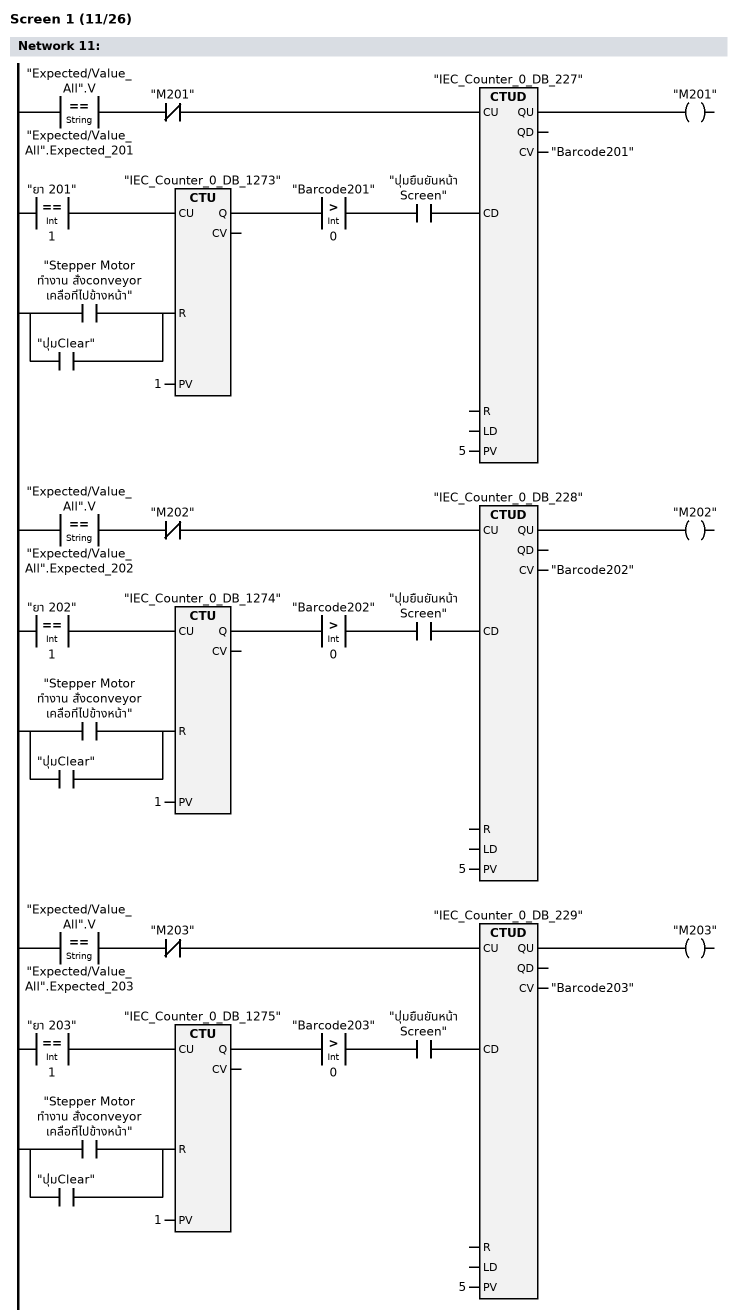
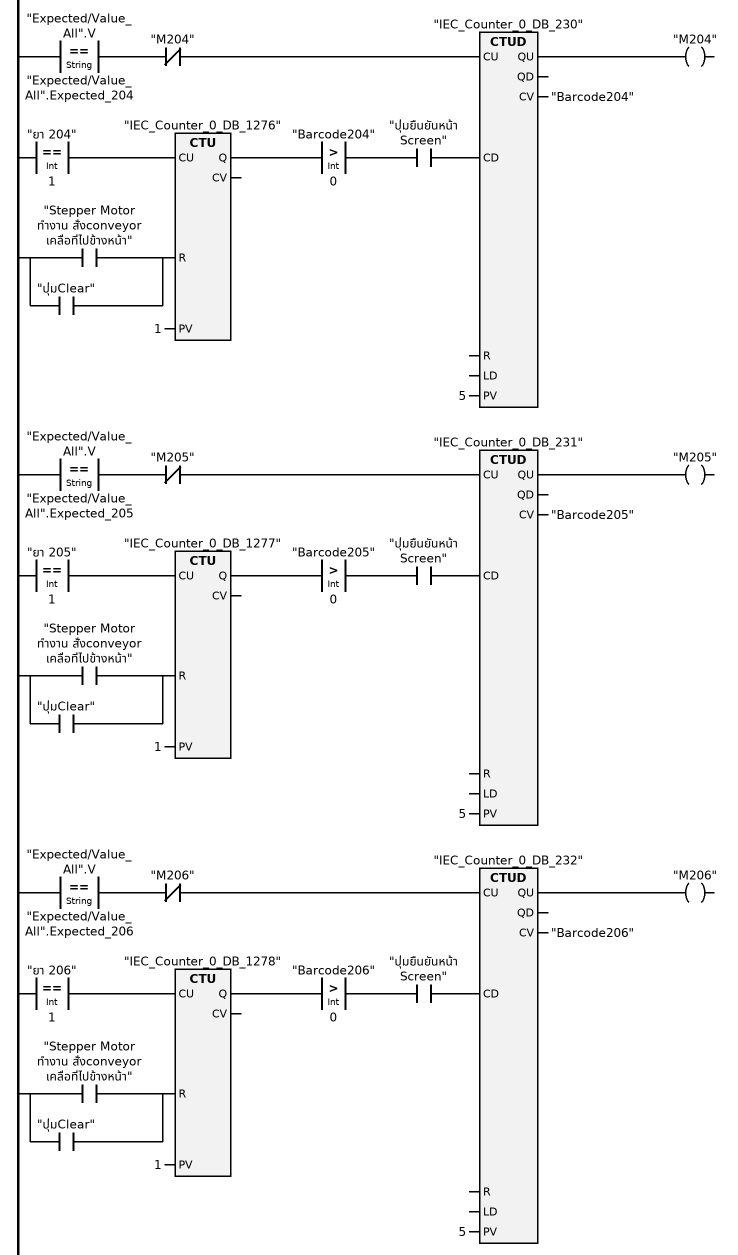
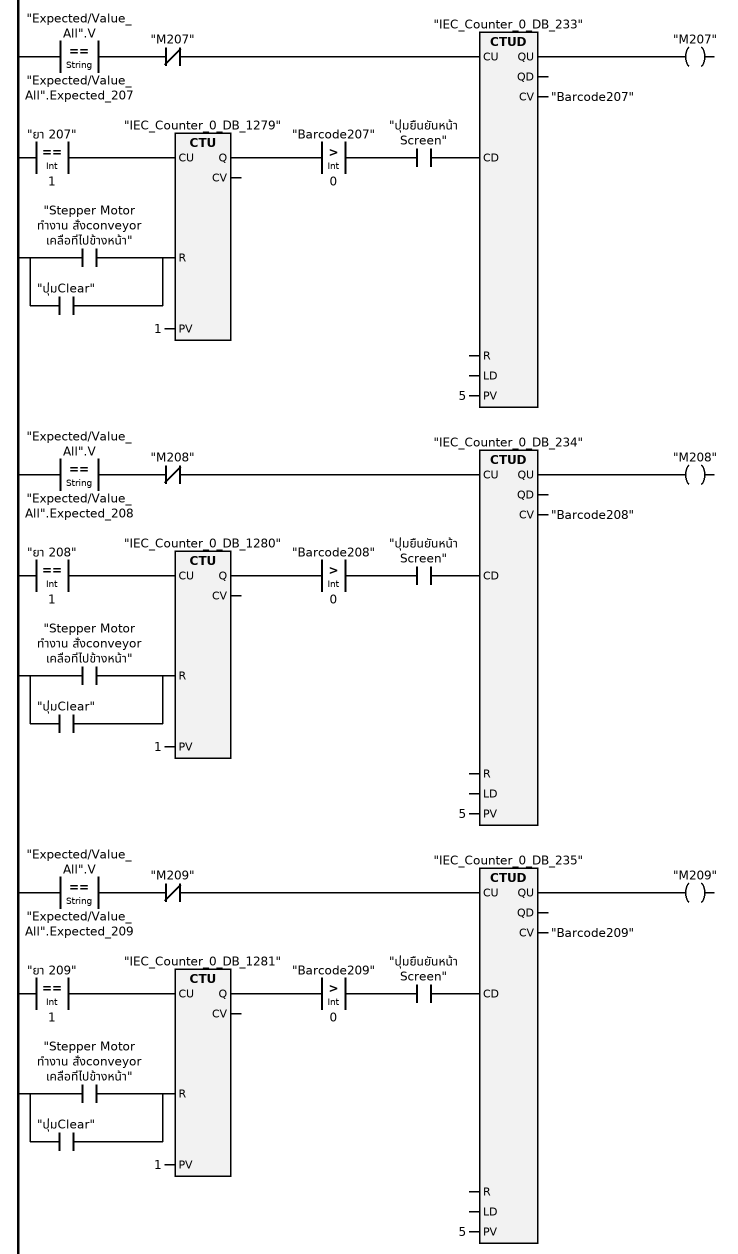
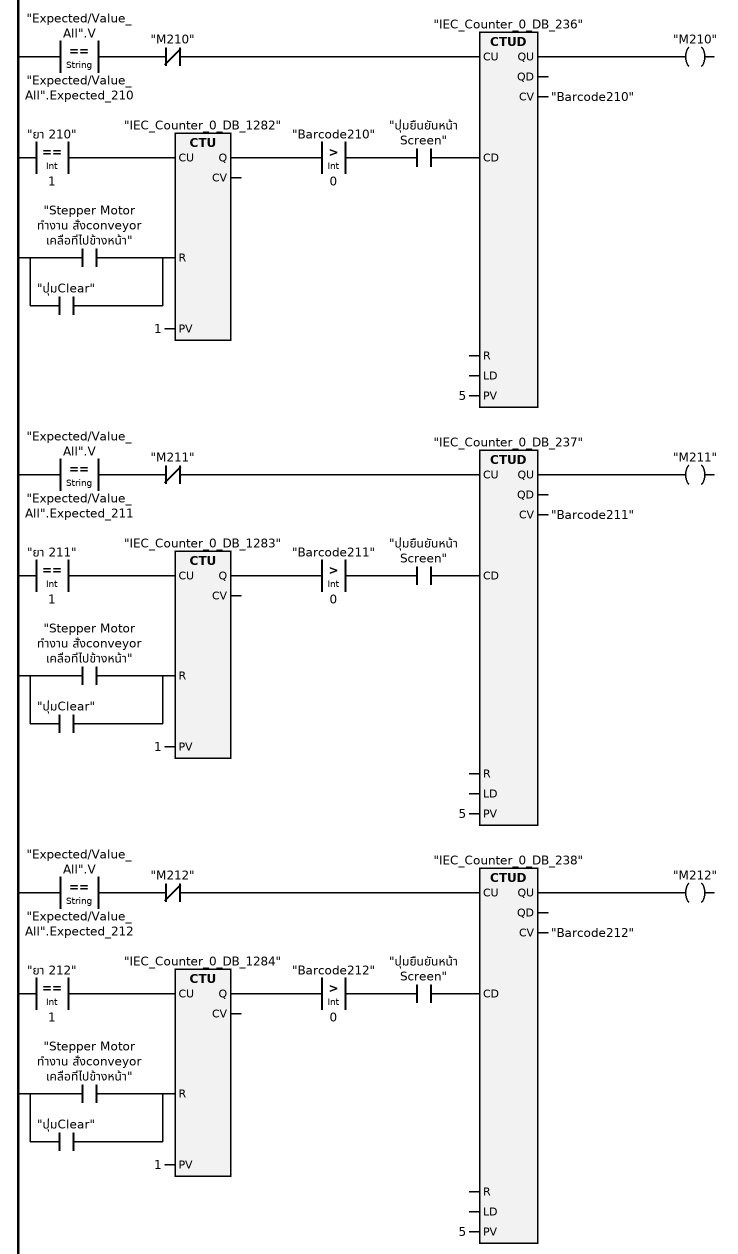
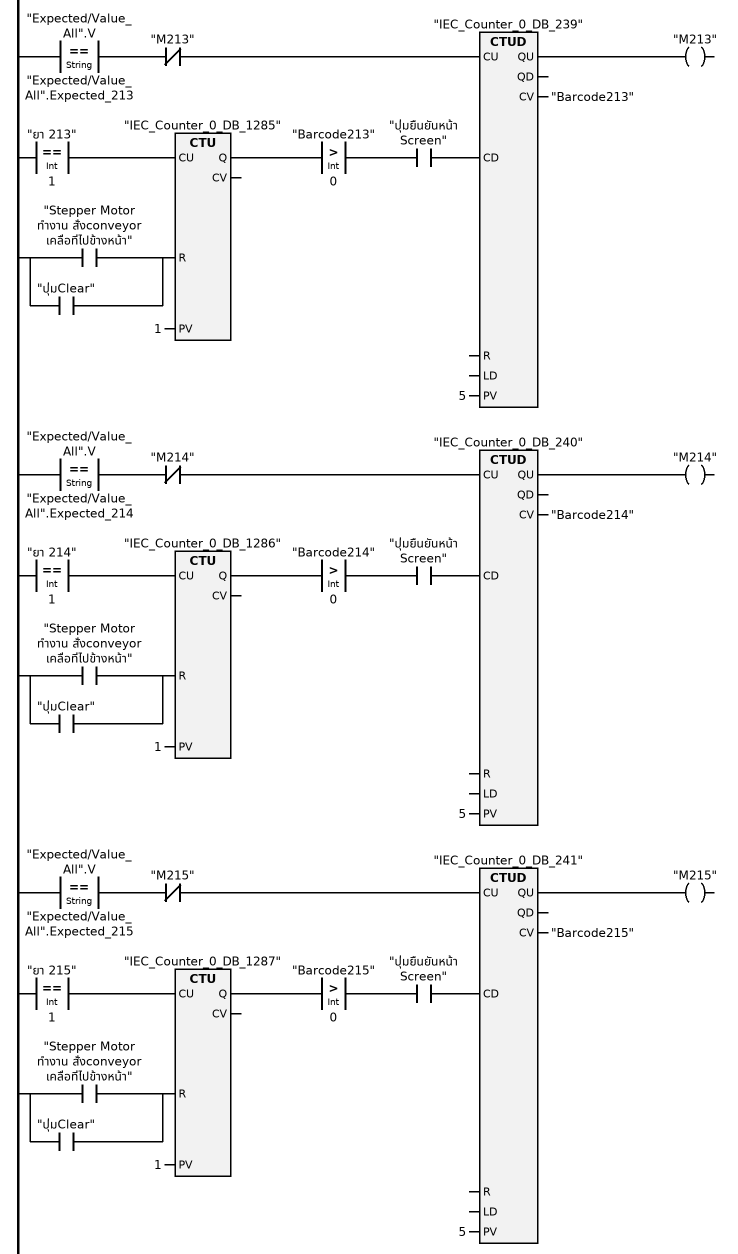
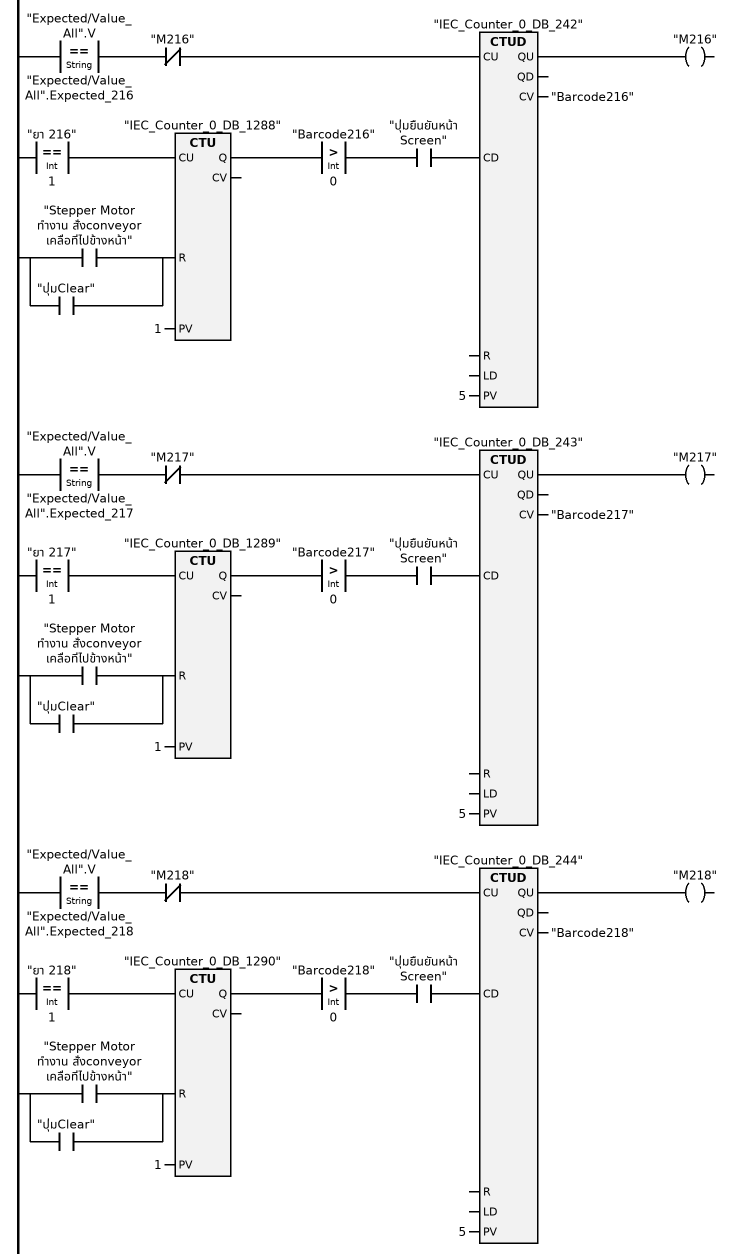
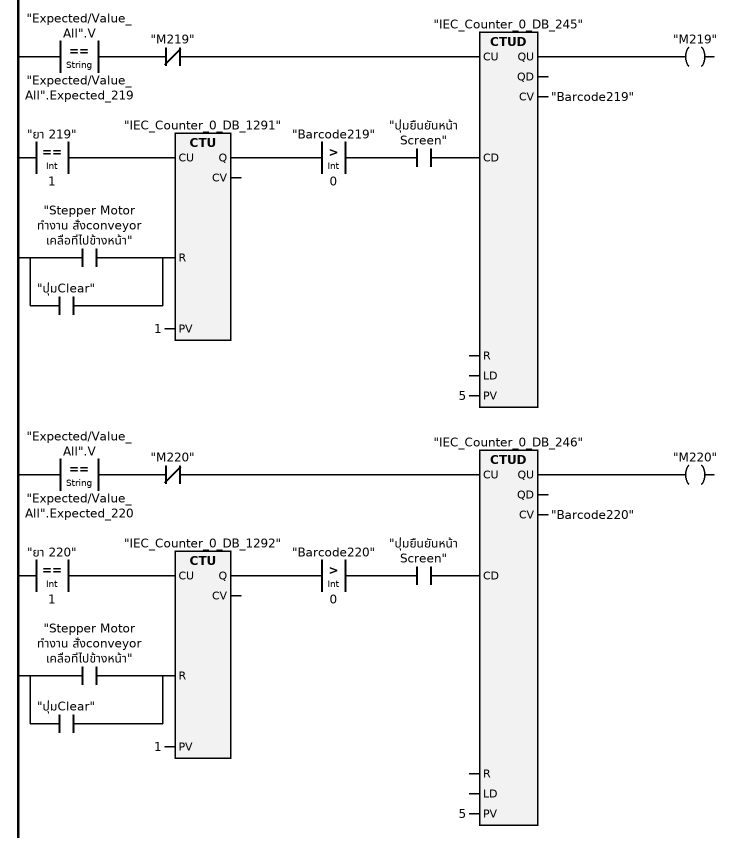
   "IEC_Counter_0_DB_1273".CTU(CU := "ยา 201" = 1,
                           R := "Stepper Motor ทำงาน สั่งconveyor เคลื่อที่ไปข้างหน้า" OR "ปุ่มClear",
                           PV := 1);
   "IEC_Counter_0_DB_227".CTUD(CU := ("Expected/Value_All".V = "Expected/Value_All".Expected_201) AND NOT "M201",
                           CD := "IEC_Counter_0_DB_1273".Q AND ("Barcode201" > 0) AND "ปุ่มยืนยันหน้า Screen",
                           PV := 5,
                           CV => "Barcode201");
   "M201" := "IEC_Counter_0_DB_227".QU;
   "IEC_Counter_0_DB_1274".CTU(CU := "ยา 202" = 1,
                           R := "Stepper Motor ทำงาน สั่งconveyor เคลื่อที่ไปข้างหน้า" OR "ปุ่มClear",
                           PV := 1);
   "IEC_Counter_0_DB_228".CTUD(CU := ("Expected/Value_All".V = "Expected/Value_All".Expected_202) AND NOT "M202",
                           CD := "IEC_Counter_0_DB_1274".Q AND ("Barcode202" > 0) AND "ปุ่มยืนยันหน้า Screen",
                           PV := 5,
                           CV => "Barcode202");
   "M202" := "IEC_Counter_0_DB_228".QU;
   "IEC_Counter_0_DB_1275".CTU(CU := "ยา 203" = 1,
                           R := "Stepper Motor ทำงาน สั่งconveyor เคลื่อที่ไปข้างหน้า" OR "ปุ่มClear",
                           PV := 1);
   "IEC_Counter_0_DB_229".CTUD(CU := ("Expected/Value_All".V = "Expected/Value_All".Expected_203) AND NOT "M203",
                           CD := "IEC_Counter_0_DB_1275".Q AND ("Barcode203" > 0) AND "ปุ่มยืนยันหน้า Screen",
                           PV := 5,
                           CV => "Barcode203");
   "M203" := "IEC_Counter_0_DB_229".QU;
   "IEC_Counter_0_DB_1276".CTU(CU := "ยา 204" = 1,
                           R := "Stepper Motor ทำงาน สั่งconveyor เคลื่อที่ไปข้างหน้า" OR "ปุ่มClear",
                           PV := 1);
   "IEC_Counter_0_DB_230".CTUD(CU := ("Expected/Value_All".V = "Expected/Value_All".Expected_204) AND NOT "M204",
                           CD := "IEC_Counter_0_DB_1276".Q AND ("Barcode204" > 0) AND "ปุ่มยืนยันหน้า Screen",
                           PV := 5,
                           CV => "Barcode204");
   "M204" := "IEC_Counter_0_DB_230".QU;
   "IEC_Counter_0_DB_1277".CTU(CU := "ยา 205" = 1,
                           R := "Stepper Motor ทำงาน สั่งconveyor เคลื่อที่ไปข้างหน้า" OR "ปุ่มClear",
                           PV := 1);
   "IEC_Counter_0_DB_231".CTUD(CU := ("Expected/Value_All".V = "Expected/Value_All".Expected_205) AND NOT "M205",
                           CD := "IEC_Counter_0_DB_1277".Q AND ("Barcode205" > 0) AND "ปุ่มยืนยันหน้า Screen",
                           PV := 5,
                           CV => "Barcode205");
   "M205" := "IEC_Counter_0_DB_231".QU;
   "IEC_Counter_0_DB_1278".CTU(CU := "ยา 206" = 1,
                           R := "Stepper Motor ทำงาน สั่งconveyor เคลื่อที่ไปข้างหน้า" OR "ปุ่มClear",
                           PV := 1);
   "IEC_Counter_0_DB_232".CTUD(CU := ("Expected/Value_All".V = "Expected/Value_All".Expected_206) AND NOT "M206",
                           CD := "IEC_Counter_0_DB_1278".Q AND ("Barcode206" > 0) AND "ปุ่มยืนยันหน้า Screen",
                           PV := 5,
                           CV => "Barcode206");
   "M206" := "IEC_Counter_0_DB_232".QU;
   "IEC_Counter_0_DB_1279".CTU(CU := "ยา 207" = 1,
                           R := "Stepper Motor ทำงาน สั่งconveyor เคลื่อที่ไปข้างหน้า" OR "ปุ่มClear",
                           PV := 1);
   "IEC_Counter_0_DB_233".CTUD(CU := ("Expected/Value_All".V = "Expected/Value_All".Expected_207) AND NOT "M207",
                           CD := "IEC_Counter_0_DB_1279".Q AND ("Barcode207" > 0) AND "ปุ่มยืนยันหน้า Screen",
                           PV := 5,
                           CV => "Barcode207");
   "M207" := "IEC_Counter_0_DB_233".QU;
   "IEC_Counter_0_DB_1280".CTU(CU := "ยา 208" = 1,
                           R := "Stepper Motor ทำงาน สั่งconveyor เคลื่อที่ไปข้างหน้า" OR "ปุ่มClear",
                           PV := 1);
   "IEC_Counter_0_DB_234".CTUD(CU := ("Expected/Value_All".V = "Expected/Value_All".Expected_208) AND NOT "M208",
                           CD := "IEC_Counter_0_DB_1280".Q AND ("Barcode208" > 0) AND "ปุ่มยืนยันหน้า Screen",
                           PV := 5,
                           CV => "Barcode208");
   "M208" := "IEC_Counter_0_DB_234".QU;
   "IEC_Counter_0_DB_1281".CTU(CU := "ยา 209" = 1,
                           R := "Stepper Motor ทำงาน สั่งconveyor เคลื่อที่ไปข้างหน้า" OR "ปุ่มClear",
                           PV := 1);
   "IEC_Counter_0_DB_235".CTUD(CU := ("Expected/Value_All".V = "Expected/Value_All".Expected_209) AND NOT "M209",
                           CD := "IEC_Counter_0_DB_1281".Q AND ("Barcode209" > 0) AND "ปุ่มยืนยันหน้า Screen",
                           PV := 5,
                           CV => "Barcode209");
   "M209" := "IEC_Counter_0_DB_235".QU;
   "IEC_Counter_0_DB_1282".CTU(CU := "ยา 210" = 1,
                           R := "Stepper Motor ทำงาน สั่งconveyor เคลื่อที่ไปข้างหน้า" OR "ปุ่มClear",
                           PV := 1);
   "IEC_Counter_0_DB_236".CTUD(CU := ("Expected/Value_All".V = "Expected/Value_All".Expected_210) AND NOT "M210",
                           CD := "IEC_Counter_0_DB_1282".Q AND ("Barcode210" > 0) AND "ปุ่มยืนยันหน้า Screen",
                           PV := 5,
                           CV => "Barcode210");
   "M210" := "IEC_Counter_0_DB_236".QU;
   "IEC_Counter_0_DB_1283".CTU(CU := "ยา 211" = 1,
                           R := "Stepper Motor ทำงาน สั่งconveyor เคลื่อที่ไปข้างหน้า" OR "ปุ่มClear",
                           PV := 1);
   "IEC_Counter_0_DB_237".CTUD(CU := ("Expected/Value_All".V = "Expected/Value_All".Expected_211) AND NOT "M211",
                           CD := "IEC_Counter_0_DB_1283".Q AND ("Barcode211" > 0) AND "ปุ่มยืนยันหน้า Screen",
                           PV := 5,
                           CV => "Barcode211");
   "M211" := "IEC_Counter_0_DB_237".QU;
   "IEC_Counter_0_DB_1284".CTU(CU := "ยา 212" = 1,
                           R := "Stepper Motor ทำงาน สั่งconveyor เคลื่อที่ไปข้างหน้า" OR "ปุ่มClear",
                           PV := 1);
   "IEC_Counter_0_DB_238".CTUD(CU := ("Expected/Value_All".V = "Expected/Value_All".Expected_212) AND NOT "M212",
                           CD := "IEC_Counter_0_DB_1284".Q AND ("Barcode212" > 0) AND "ปุ่มยืนยันหน้า Screen",
                           PV := 5,
                           CV => "Barcode212");
   "M212" := "IEC_Counter_0_DB_238".QU;
   "IEC_Counter_0_DB_1285".CTU(CU := "ยา 213" = 1,
                           R := "Stepper Motor ทำงาน สั่งconveyor เคลื่อที่ไปข้างหน้า" OR "ปุ่มClear",
                           PV := 1);
   "IEC_Counter_0_DB_239".CTUD(CU := ("Expected/Value_All".V = "Expected/Value_All".Expected_213) AND NOT "M213",
                           CD := "IEC_Counter_0_DB_1285".Q AND ("Barcode213" > 0) AND "ปุ่มยืนยันหน้า Screen",
                           PV := 5,
                           CV => "Barcode213");
   "M213" := "IEC_Counter_0_DB_239".QU;
   "IEC_Counter_0_DB_1286".CTU(CU := "ยา 214" = 1,
                           R := "Stepper Motor ทำงาน สั่งconveyor เคลื่อที่ไปข้างหน้า" OR "ปุ่มClear",
                           PV := 1);
   "IEC_Counter_0_DB_240".CTUD(CU := ("Expected/Value_All".V = "Expected/Value_All".Expected_214) AND NOT "M214",
                           CD := "IEC_Counter_0_DB_1286".Q AND ("Barcode214" > 0) AND "ปุ่มยืนยันหน้า Screen",
                           PV := 5,
                           CV => "Barcode214");
   "M214" := "IEC_Counter_0_DB_240".QU;
   "IEC_Counter_0_DB_1287".CTU(CU := "ยา 215" = 1,
                           R := "Stepper Motor ทำงาน สั่งconveyor เคลื่อที่ไปข้างหน้า" OR "ปุ่มClear",
                           PV := 1);
   "IEC_Counter_0_DB_241".CTUD(CU := ("Expected/Value_All".V = "Expected/Value_All".Expected_215) AND NOT "M215",
                           CD := "IEC_Counter_0_DB_1287".Q AND ("Barcode215" > 0) AND "ปุ่มยืนยันหน้า Screen",
                           PV := 5,
                           CV => "Barcode215");
   "M215" := "IEC_Counter_0_DB_241".QU;
   "IEC_Counter_0_DB_1288".CTU(CU := "ยา 216" = 1,
                           R := "Stepper Motor ทำงาน สั่งconveyor เคลื่อที่ไปข้างหน้า" OR "ปุ่มClear",
                           PV := 1);
   "IEC_Counter_0_DB_242".CTUD(CU := ("Expected/Value_All".V = "Expected/Value_All".Expected_216) AND NOT "M216",
                           CD := "IEC_Counter_0_DB_1288".Q AND ("Barcode216" > 0) AND "ปุ่มยืนยันหน้า Screen",
                           PV := 5,
                           CV => "Barcode216");
   "M216" := "IEC_Counter_0_DB_242".QU;
   "IEC_Counter_0_DB_1289".CTU(CU := "ยา 217" = 1,
                           R := "Stepper Motor ทำงาน สั่งconveyor เคลื่อที่ไปข้างหน้า" OR "ปุ่มClear",
                           PV := 1);
   "IEC_Counter_0_DB_243".CTUD(CU := ("Expected/Value_All".V = "Expected/Value_All".Expected_217) AND NOT "M217",
                           CD := "IEC_Counter_0_DB_1289".Q AND ("Barcode217" > 0) AND "ปุ่มยืนยันหน้า Screen",
                           PV := 5,
                           CV => "Barcode217");
   "M217" := "IEC_Counter_0_DB_243".QU;
   "IEC_Counter_0_DB_1290".CTU(CU := "ยา 218" = 1,
                           R := "Stepper Motor ทำงาน สั่งconveyor เคลื่อที่ไปข้างหน้า" OR "ปุ่มClear",
                           PV := 1);
   "IEC_Counter_0_DB_244".CTUD(CU := ("Expected/Value_All".V = "Expected/Value_All".Expected_218) AND NOT "M218",
                           CD := "IEC_Counter_0_DB_1290".Q AND ("Barcode218" > 0) AND "ปุ่มยืนยันหน้า Screen",
                           PV := 5,
                           CV => "Barcode218");
   "M218" := "IEC_Counter_0_DB_244".QU;
   "IEC_Counter_0_DB_1291".CTU(CU := "ยา 219" = 1,
                           R := "Stepper Motor ทำงาน สั่งconveyor เคลื่อที่ไปข้างหน้า" OR "ปุ่มClear",
                           PV := 1);
   "IEC_Counter_0_DB_245".CTUD(CU := ("Expected/Value_All".V = "Expected/Value_All".Expected_219) AND NOT "M219",
                           CD := "IEC_Counter_0_DB_1291".Q AND ("Barcode219" > 0) AND "ปุ่มยืนยันหน้า Screen",
                           PV := 5,
                           CV => "Barcode219");
   "M219" := "IEC_Counter_0_DB_245".QU;
   "IEC_Counter_0_DB_1292".CTU(CU := "ยา 220" = 1,
                           R := "Stepper Motor ทำงาน สั่งconveyor เคลื่อที่ไปข้างหน้า" OR "ปุ่มClear",
                           PV := 1);
   "IEC_Counter_0_DB_246".CTUD(CU := ("Expected/Value_All".V = "Expected/Value_All".Expected_220) AND NOT "M220",
                           CD := "IEC_Counter_0_DB_1292".Q AND ("Barcode220" > 0) AND "ปุ่มยืนยันหน้า Screen",
                           PV := 5,
                           CV => "Barcode220");
   "M220" := "IEC_Counter_0_DB_246".QU;
END_REGION

REGION Network 12
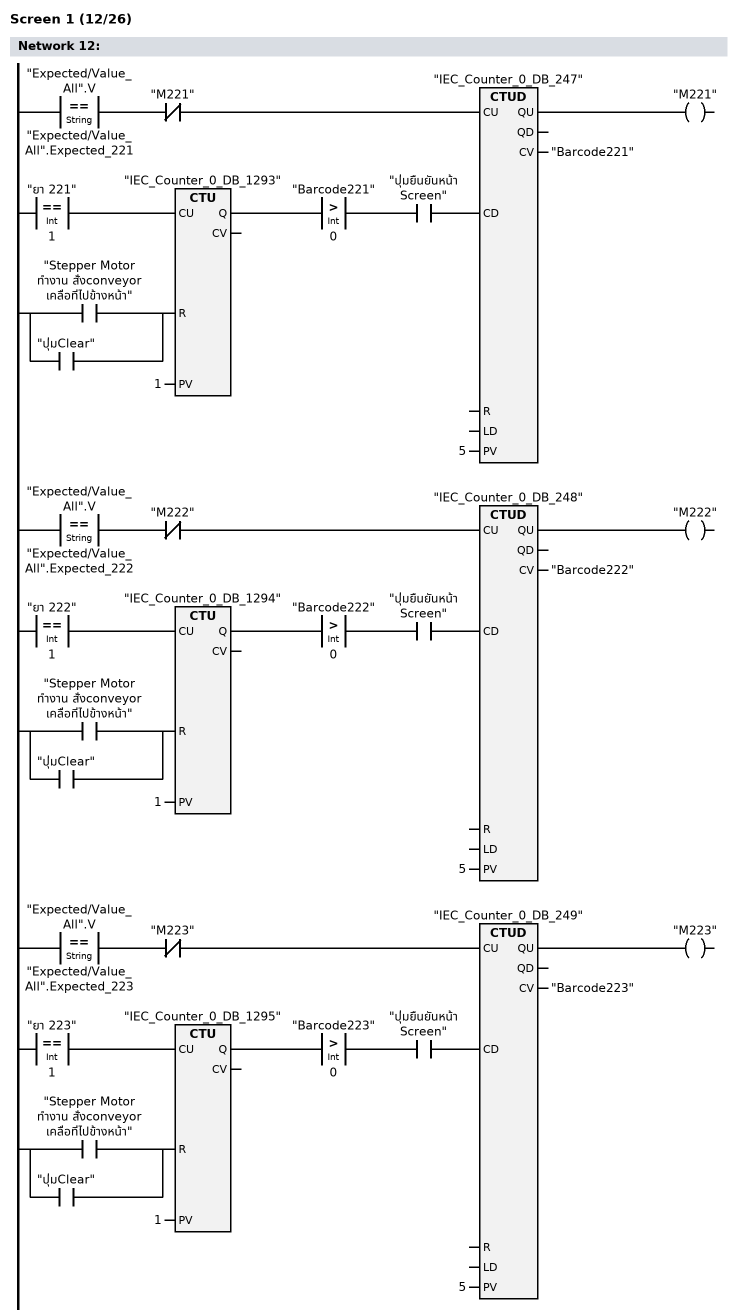
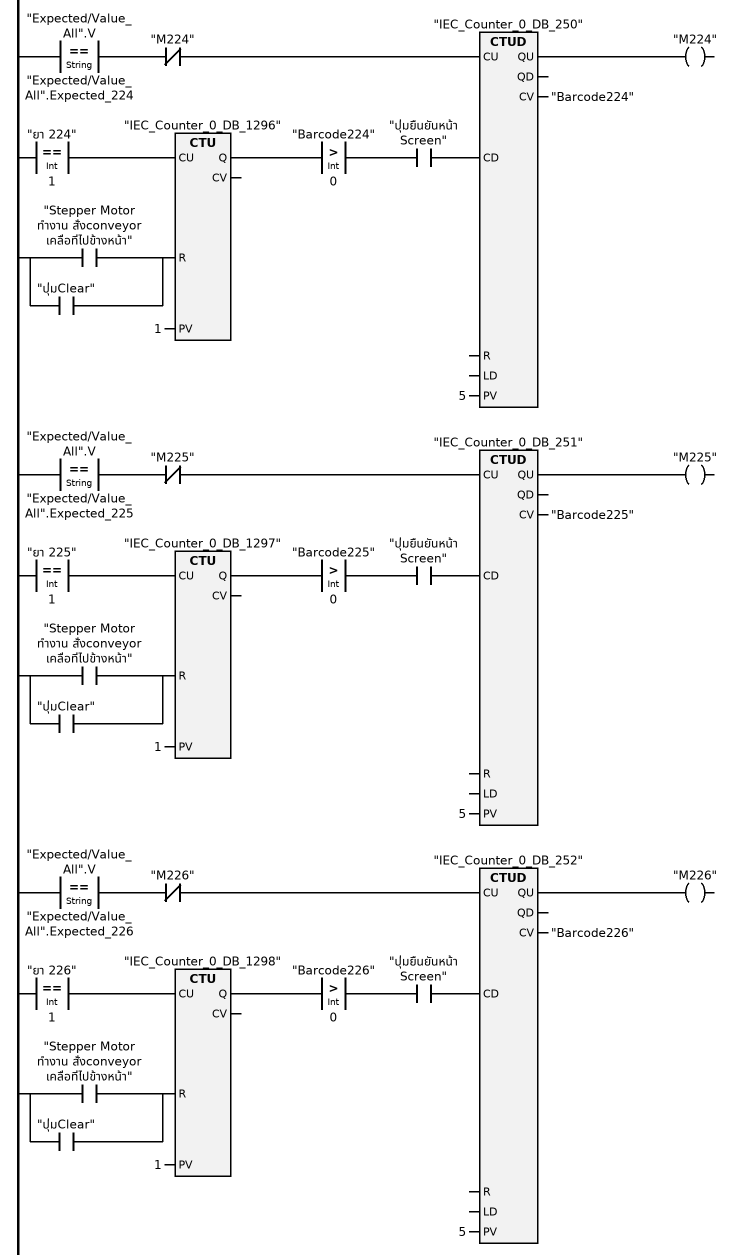
